(* IEC 61131-3 sources: TetherPLC/compat/tc3 (part 4) *)

(* ---- tc3_mcpath.st ---- *)
// Tc3_McCoordinatedMotion — MC path preparation + execution
// (TF5410 collision-avoidance / coordinated-motion bundle).
//
// This tranche implements the linear/dwell path subset:
//   MC_MoveLinearAbsolutePreparation, MC_MoveDirectPreparation
//   (flattened alias of the linear absolute segment),
//   MC_DwellTimePreparation, MC_MovePath.
// Path objects live in the tplc-path service via the FB_Path
// builtin; group membership comes from FB_McGroup.  Circular,
// blending and blocker segment types, MC_CalcTrafo, the CA move
// family, track following and compensation remain deferred.
//
// Flattened types (the ST dialect has no STRUCT/POINTER/REFERENCE
// support):
//   MC_PATH_DATA_REF     -> PathData : UDINT path handle (1..8)
//   Position (POINTER TO LREAL array) -> Position : ARRAY[0..15]
//                            OF LREAL + PositionCount
//   DwellTime (TIME)     -> DwellTime : UDINT milliseconds
//   BufferMode           -> UDINT (accepted, buffered queuing not
//                            modeled: every Execute edge appends a
//                            segment immediately)
//   AXES_GROUP_REF       -> AxesGroup : UDINT group handle
//
// Semantics:
//   * Preparation FBs append one segment on the Execute rising
//     edge. Linear segments store absolute user-unit positions and
//     trapezoid limits (Velocity/Acceleration; Deceleration and
//     Jerk are accepted but the service uses Acceleration for both
//     ramps). Dwell segments hold position for DwellTime ms.
//   * MC_MovePath on Execute captures each member axis's current
//     position (0x6064) as the path start, switches every member
//     to CSP mode (0x6060=8), then streams interpolated 0x607A
//     targets each scan until the path duration elapses. Positions
//     are interpolated in path parameter space on the dominant
//     axis, so all axes arrive together (coordinated motion).
//   * Segment targets chain: segment k starts where segment k-1
//     ended; the first segment starts at the captured positions.
//   * Busy stays TRUE while the path runs; Done pulses for one
//     scan at path end; Error carries service/axis failures.

// ---- shared path helper: ensure a valid PathData handle ----
// Returns TRUE and leaves `h` set to a usable path handle, or
// FALSE when the service table is full.

FUNCTION_BLOCK MC_MoveLinearAbsolutePreparation
VAR_INPUT
    Execute : BOOL;
    Position : ARRAY[0..15] OF LREAL;
    PositionCount : UDINT;
    Velocity : LREAL;
    Acceleration : LREAL;
    Deceleration : LREAL := 0.0;
    Jerk : LREAL := 0.0;
    BufferMode : UDINT := 1;
END_VAR
VAR_IN_OUT
    PathData : UDINT;
END_VAR
VAR_OUTPUT
    Error : BOOL;
    ErrorId : UDINT;
END_VAR
VAR
    p : FB_Path;
    exPrev : BOOL;
    edge : BOOL;
    i : UDINT;
END_VAR
edge := Execute AND NOT exPrev; exPrev := Execute;
Error := FALSE; ErrorId := 0;
IF edge THEN
    p.HANDLE := PathData;
    IF PathData = 0 THEN
        p.OP := 0; p();
        IF p.STATUS = 0 THEN PathData := p.HANDLE; END_IF;
    END_IF;
    IF PathData <> 0 AND PositionCount >= 1 AND
       PositionCount <= 16 THEN
        FOR i := 0 TO 15 DO p.POS[i] := Position[i]; END_FOR;
        p.OP := 2; p.AUX := 1; p.AUX2 := PositionCount;
        p.F1 := Velocity; p.F2 := Acceleration; p.F3 := 0.0;
        p.HANDLE := PathData; p();
        IF p.STATUS <> 0 THEN
            Error := TRUE;
            IF p.STATUS < 0 THEN ErrorId := 0 - p.STATUS; END_IF;
        END_IF;
    ELSE
        Error := TRUE; ErrorId := 16#4D01;
    END_IF;
END_IF;
END_FUNCTION_BLOCK

// MC_MoveDirectPreparation: TwinCAT "direct" segments are absolute
// linear moves without blending lookahead.  Flattened to the same
// linear segment; BufferMode is accepted for signature parity.
FUNCTION_BLOCK MC_MoveDirectPreparation
VAR_INPUT
    Execute : BOOL;
    Position : ARRAY[0..15] OF LREAL;
    PositionCount : UDINT;
    Velocity : LREAL;
    Acceleration : LREAL;
    Deceleration : LREAL := 0.0;
    Jerk : LREAL := 0.0;
    BufferMode : UDINT := 1;
END_VAR
VAR_IN_OUT
    PathData : UDINT;
END_VAR
VAR_OUTPUT
    Error : BOOL;
    ErrorId : UDINT;
END_VAR
VAR
    p : FB_Path;
    exPrev : BOOL;
    edge : BOOL;
    i : UDINT;
END_VAR
edge := Execute AND NOT exPrev; exPrev := Execute;
Error := FALSE; ErrorId := 0;
IF edge THEN
    p.HANDLE := PathData;
    IF PathData = 0 THEN
        p.OP := 0; p();
        IF p.STATUS = 0 THEN PathData := p.HANDLE; END_IF;
    END_IF;
    IF PathData <> 0 AND PositionCount >= 1 AND
       PositionCount <= 16 THEN
        FOR i := 0 TO 15 DO p.POS[i] := Position[i]; END_FOR;
        p.OP := 2; p.AUX := 1; p.AUX2 := PositionCount;
        p.F1 := Velocity; p.F2 := Acceleration; p.F3 := 0.0;
        p.HANDLE := PathData; p();
        IF p.STATUS <> 0 THEN
            Error := TRUE;
            IF p.STATUS < 0 THEN ErrorId := 0 - p.STATUS; END_IF;
        END_IF;
    ELSE
        Error := TRUE; ErrorId := 16#4D01;
    END_IF;
END_IF;
END_FUNCTION_BLOCK

FUNCTION_BLOCK MC_DwellTimePreparation
VAR_INPUT
    Execute : BOOL;
    DwellTime : UDINT;   // milliseconds (TIME flattened)
    BufferMode : UDINT := 1;
END_VAR
VAR_IN_OUT
    PathData : UDINT;
END_VAR
VAR_OUTPUT
    Error : BOOL;
    ErrorId : UDINT;
END_VAR
VAR
    p : FB_Path;
    exPrev : BOOL;
    edge : BOOL;
END_VAR
edge := Execute AND NOT exPrev; exPrev := Execute;
Error := FALSE; ErrorId := 0;
IF edge THEN
    p.HANDLE := PathData;
    IF PathData = 0 THEN
        p.OP := 0; p();
        IF p.STATUS = 0 THEN PathData := p.HANDLE; END_IF;
    END_IF;
    IF PathData <> 0 THEN
        p.OP := 2; p.AUX := 3; p.AUX2 := 0;
        p.F1 := 0.0; p.F2 := 0.0; p.F3 := DwellTime;
        p.HANDLE := PathData; p();
        IF p.STATUS <> 0 THEN
            Error := TRUE;
            IF p.STATUS < 0 THEN ErrorId := 0 - p.STATUS; END_IF;
        END_IF;
    ELSE
        Error := TRUE; ErrorId := 16#4D01;
    END_IF;
END_IF;
END_FUNCTION_BLOCK

FUNCTION_BLOCK MC_MovePath
VAR_INPUT
    Execute : BOOL;
END_VAR
VAR_IN_OUT
    AxesGroup : UDINT;
    PathData : UDINT;
END_VAR
VAR_OUTPUT
    Done : BOOL;
    Busy : BOOL;
    CommandAborted : BOOL;
    Error : BOOL;
    ErrorId : UDINT;
END_VAR
VAR
    mg : FB_McGroup;
    p : FB_Path;
    ax : FB_MotionAxis;
    exPrev : BOOL;
    exEdge : BOOL;
    active : BOOL;
    issued : BOOL;
    t0 : LREAL;
    pathT : LREAL;
    lastNow : LREAL;
    blkWait : BOOL;
    trafoGen : UDINT;
    lastTrafoGen : UDINT;
    dn : LREAL;
    i : UDINT;
    n : UDINT;
    axh : UDINT;
    startPos : ARRAY[0..15] OF LREAL;
END_VAR
mg.GRP := AxesGroup;
mg.OP := 10; mg();
AxesGroup := mg.GRP;
n := mg.NAXES;
exEdge := Execute AND NOT exPrev; exPrev := Execute;
Done := FALSE; Busy := FALSE;
CommandAborted := FALSE; Error := FALSE; ErrorId := 0;
IF exEdge THEN
    active := TRUE; issued := FALSE;
END_IF;
IF active THEN
    IF NOT issued THEN
        /* capture current positions as the path start */
        FOR i := 0 TO 15 DO
            startPos[i] := 0.0;
            IF i < n THEN
                axh := mg.AXES[i];
                ax.AXIS := axh; ax.OP := 4; ax.INDEX := 16#6064; ax();
                startPos[i] := DINT_TO_LREAL(ax.VALUE);
            END_IF;
        END_FOR;
        FOR i := 0 TO 15 DO p.POS[i] := startPos[i]; END_FOR;
        p.OP := 3; p.AUX := n; p.HANDLE := PathData; p();
        IF p.STATUS <> 0 THEN
            Error := TRUE;
            IF p.STATUS < 0 THEN ErrorId := 0 - p.STATUS; END_IF;
            active := FALSE;
        ELSE
            PathData := p.HANDLE;
            /* bind the path to the group for trajectory readback */
            p.OP := 9; p.AUX := AxesGroup; p.HANDLE := PathData; p();
            t0 := p.NOW;
            pathT := 0.0; lastNow := p.NOW;
            /* switch members to CSP mode for 0x607A streaming */
            FOR i := 0 TO 15 DO
                IF i < n THEN
                    axh := mg.AXES[i];
                    ax.AXIS := axh; ax.OP := 5;
                    ax.INDEX := 16#6060; ax.VALUE := 8; ax();
                END_IF;
            END_FOR;
            issued := TRUE;
        END_IF;
    END_IF;
    IF issued THEN
        /* blocker query freezes path time while the path is held
           at an unreleased blocker gate */
        p.OP := 7; p.HANDLE := PathData; p();
        blkWait := p.AUX = 1;
        dn := p.NOW - lastNow; lastNow := p.NOW;
        IF NOT blkWait THEN pathT := pathT + dn; END_IF;
        /* apply pending coordinate-transform markers: the service
           bumps AUX2 whenever the pending id changes */
        p.OP := 11; p.HANDLE := PathData; p();
        trafoGen := p.AUX2;
        IF trafoGen <> lastTrafoGen AND p.F1 <> 0.0 THEN
            lastTrafoGen := trafoGen;
            mg.OP := 9; mg.COORD := LREAL_TO_DINT(p.F1); mg();
        END_IF;
        p.OP := 4; p.F1 := pathT; p.HANDLE := PathData; p();
        IF p.STATUS <> 0 THEN
            Error := TRUE;
            IF p.STATUS < 0 THEN ErrorId := 0 - p.STATUS; END_IF;
            active := FALSE; CommandAborted := TRUE;
        ELSE
            FOR i := 0 TO 15 DO
                IF i < n THEN
                    axh := mg.AXES[i];
                    ax.AXIS := axh; ax.OP := 5;
                    ax.INDEX := 16#607A;
                    ax.VALUE := LREAL_TO_DINT(p.POS[i]); ax();
                END_IF;
            END_FOR;
            IF p.DONE = 1 THEN
                Done := TRUE; active := FALSE;
            END_IF;
        END_IF;
    END_IF;
    Busy := active;
END_IF;
END_FUNCTION_BLOCK

// MC_MoveCircularAbsolutePreparation: appends a circular segment.
// CircMode flattens MC_CIRC_MODE (1=mcCircModeCenter: AuxPoint is
// the circle center and must be equidistant from start/end;
// 2=mcCircModeBorder: AuxPoint lies on the circle). The circle is
// evaluated in the plane of position entries 0/1; entries >=2
// interpolate linearly. PathChoice: 1=counter-clockwise,
// 2=clockwise. TransitionMode/TransitionParameter/InvokeId/
// DynamicConstraints are accepted for signature parity but not
// modeled.
FUNCTION_BLOCK MC_MoveCircularAbsolutePreparation
VAR_INPUT
    Execute : BOOL;
    CircMode : UDINT;
    AuxPoint : ARRAY[0..15] OF LREAL;
    AuxPointCount : UDINT;
    EndPoint : ARRAY[0..15] OF LREAL;
    EndPointCount : UDINT;
    PathChoice : UDINT := 1;
    Velocity : LREAL;
    Acceleration : LREAL;
    Deceleration : LREAL := 0.0;
    Jerk : LREAL := 0.0;
    BufferMode : UDINT := 1;
    TransitionMode : UDINT := 0;
    TransitionParameter : ARRAY[0..15] OF LREAL;
    TransitionParameterCount : UDINT := 0;
    InvokeId : UDINT := 0;
END_VAR
VAR_IN_OUT
    PathData : UDINT;
END_VAR
VAR_OUTPUT
    Error : BOOL;
    ErrorId : UDINT;
END_VAR
VAR
    p : FB_Path;
    exPrev : BOOL;
    edge : BOOL;
    i : UDINT;
END_VAR
edge := Execute AND NOT exPrev; exPrev := Execute;
Error := FALSE; ErrorId := 0;
IF edge THEN
    p.HANDLE := PathData;
    IF PathData = 0 THEN
        p.OP := 0; p();
        IF p.STATUS = 0 THEN PathData := p.HANDLE; END_IF;
    END_IF;
    IF PathData <> 0 AND EndPointCount >= 1 AND EndPointCount <= 16
       AND CircMode >= 1 AND CircMode <= 2 THEN
        FOR i := 0 TO 15 DO
            p.POS[i] := EndPoint[i];
            p.AUXP[i] := AuxPoint[i];
        END_FOR;
        p.OP := 6; p.AUX := CircMode; p.FLAGS := AuxPointCount;
        p.AUX2 := EndPointCount; p.F3 := PathChoice;
        p.F1 := Velocity; p.F2 := Acceleration;
        p.HANDLE := PathData; p();
        IF p.STATUS <> 0 THEN
            Error := TRUE;
            IF p.STATUS < 0 THEN ErrorId := 0 - p.STATUS; END_IF;
        END_IF;
    ELSE
        Error := TRUE; ErrorId := 16#4D01;
    END_IF;
END_IF;
END_FUNCTION_BLOCK

// MC_MoveBlendingPreparation: appends a junction transition segment.
// TwinCAT uses it to program velocity blending between segments;
// this implementation holds the path end position for
// TransitionParameter[0] milliseconds (real corner-cutting/lookahead
// blending is not modeled — documented deviation). Velocity/
// Acceleration/Deceleration/Jerk are accepted for signature parity.
FUNCTION_BLOCK MC_MoveBlendingPreparation
VAR_INPUT
    Execute : BOOL;
    Velocity : LREAL;
    Acceleration : LREAL;
    Deceleration : LREAL := 0.0;
    Jerk : LREAL := 0.0;
    BufferMode : UDINT := 1;
    TransitionMode : UDINT := 0;
    TransitionParameter : ARRAY[0..15] OF LREAL;
    TransitionParameterCount : UDINT := 0;
    InvokeId : UDINT := 0;
END_VAR
VAR_IN_OUT
    PathData : UDINT;
END_VAR
VAR_OUTPUT
    Error : BOOL;
    ErrorId : UDINT;
END_VAR
VAR
    p : FB_Path;
    exPrev : BOOL;
    edge : BOOL;
END_VAR
edge := Execute AND NOT exPrev; exPrev := Execute;
Error := FALSE; ErrorId := 0;
IF edge THEN
    p.HANDLE := PathData;
    IF PathData = 0 THEN
        p.OP := 0; p();
        IF p.STATUS = 0 THEN PathData := p.HANDLE; END_IF;
    END_IF;
    IF PathData <> 0 THEN
        p.OP := 2; p.AUX := 4; p.AUX2 := 0;
        p.F1 := 0.0; p.F2 := 0.0;
        IF TransitionParameterCount >= 1 THEN
            p.F3 := TransitionParameter[0];
        ELSE
            p.F3 := 0.0;
        END_IF;
        p.HANDLE := PathData; p();
        IF p.STATUS <> 0 THEN
            Error := TRUE;
            IF p.STATUS < 0 THEN ErrorId := 0 - p.STATUS; END_IF;
        END_IF;
    ELSE
        Error := TRUE; ErrorId := 16#4D01;
    END_IF;
END_IF;
END_FUNCTION_BLOCK

// MC_BlockerPreparation: appends a blocker gate at the current path
// junction. The path holds position there during MC_MovePath until
// MC_ReleaseBlocker opens the gate. BufferMode is accepted for
// signature parity.
FUNCTION_BLOCK MC_BlockerPreparation
VAR_INPUT
    Execute : BOOL;
    BlockerId : UDINT;
    BufferMode : UDINT := 1;
END_VAR
VAR_IN_OUT
    PathData : UDINT;
END_VAR
VAR_OUTPUT
    Error : BOOL;
    ErrorId : UDINT;
END_VAR
VAR
    p : FB_Path;
    exPrev : BOOL;
    edge : BOOL;
END_VAR
edge := Execute AND NOT exPrev; exPrev := Execute;
Error := FALSE; ErrorId := 0;
IF edge THEN
    p.HANDLE := PathData;
    IF PathData = 0 THEN
        p.OP := 0; p();
        IF p.STATUS = 0 THEN PathData := p.HANDLE; END_IF;
    END_IF;
    IF PathData <> 0 AND BlockerId > 0 THEN
        p.OP := 2; p.AUX := 5; p.AUX2 := 0;
        p.F1 := 0.0; p.F2 := 0.0; p.F3 := BlockerId;
        p.HANDLE := PathData; p();
        IF p.STATUS <> 0 THEN
            Error := TRUE;
            IF p.STATUS < 0 THEN ErrorId := 0 - p.STATUS; END_IF;
        END_IF;
    ELSE
        Error := TRUE; ErrorId := 16#4D01;
    END_IF;
END_IF;
END_FUNCTION_BLOCK

// MC_ReleaseBlocker: opens every blocker gate with the given id on
// the next eval. The TwinCAT signature carries only AxesGroup; the
// flattened implementation releases by BlockerId across all path
// objects (blocker ids are user-unique per machine).
FUNCTION_BLOCK MC_ReleaseBlocker
VAR_INPUT
    Execute : BOOL;
    BlockerId : UDINT;
END_VAR
VAR_IN_OUT
    AxesGroup : UDINT;
END_VAR
VAR_OUTPUT
    Done : BOOL;
    Busy : BOOL;
    Error : BOOL;
    ErrorId : UDINT;
END_VAR
VAR
    p : FB_Path;
    mg : FB_McGroup;
    exPrev : BOOL;
    edge : BOOL;
    ok : BOOL;
END_VAR
ok := FALSE;
edge := Execute AND NOT exPrev;
mg.GRP := AxesGroup; mg.OP := 1; mg();
AxesGroup := mg.GRP;
IF edge THEN
    p.OP := 8; p.F1 := BlockerId; p();
    IF p.STATUS = 0 THEN ok := TRUE; END_IF;
END_IF;
exPrev := Execute;
Done := ok; Busy := FALSE;
Error := edge AND NOT ok;
IF edge AND p.STATUS < 0 THEN ErrorId := 0 - p.STATUS; END_IF;
END_FUNCTION_BLOCK

// MC_GroupReadBlockerStatus: reports whether the most recent path
// eval is held at an unreleased blocker. The group linkage is
// approximated — the service reports the last-evaluated path's gate
// state.
FUNCTION_BLOCK MC_GroupReadBlockerStatus
VAR_INPUT
    Enable : BOOL;
END_VAR
VAR_IN_OUT
    AxesGroup : UDINT;
END_VAR
VAR_OUTPUT
    Valid : BOOL;
    Busy : BOOL;
    Blocked : BOOL;
    BlockerId : UDINT;
    Error : BOOL;
    ErrorId : UDINT;
END_VAR
VAR
    p : FB_Path;
    mg : FB_McGroup;
END_VAR
Valid := FALSE; Busy := FALSE; Blocked := FALSE;
BlockerId := 0; Error := FALSE; ErrorId := 0;
mg.GRP := AxesGroup; mg.OP := 6; mg();
IF Enable AND mg.STATUS = 0 THEN
    Valid := TRUE;
    p.OP := 7; p();
    IF p.STATUS = 0 THEN
        Blocked := p.AUX = 1;
        BlockerId := LREAL_TO_DINT(p.F1);
    ELSE
        Error := TRUE;
        IF p.STATUS < 0 THEN ErrorId := 0 - p.STATUS; END_IF;
    END_IF;
END_IF;
END_FUNCTION_BLOCK

// MC_GroupReadTrajectoryInformation: reads the current and next
// path segments for the group the executing MC_MovePath is bound
// to. Entries flatten MC_TRAJECTORY_ENTRY: InvokeId is approximated
// by the 1-based segment index, Active marks blend/blocker
// segments, RemainingDuration is seconds and
// RemainingCartesianLength is dominant-axis user units, all as of
// the most recent path eval.
FUNCTION_BLOCK MC_GroupReadTrajectoryInformation
VAR_INPUT
    Enable : BOOL;
END_VAR
VAR_IN_OUT
    AxesGroup : UDINT;
END_VAR
VAR_OUTPUT
    Valid : BOOL;
    Busy : BOOL;
    Error : BOOL;
    ErrorId : UDINT;
    EntryCount : UDINT;
    TrajInvokeId : ARRAY[0..9] OF UDINT;
    TrajActive : ARRAY[0..9] OF BOOL;
    TrajRemLen : ARRAY[0..9] OF LREAL;
    TrajRemDur : ARRAY[0..9] OF LREAL;
END_VAR
VAR
    p : FB_Path;
    mg : FB_McGroup;
    i : UDINT;
END_VAR
Valid := FALSE; Busy := FALSE; Error := FALSE; ErrorId := 0;
EntryCount := 0;
mg.GRP := AxesGroup; mg.OP := 6; mg();
IF Enable AND mg.STATUS = 0 THEN
    Valid := TRUE;
    p.OP := 10; p.AUX := AxesGroup; p();
    IF p.STATUS = 0 THEN
        EntryCount := p.NSEG;
        FOR i := 0 TO 9 DO
            TrajInvokeId[i] := p.TRID[i];
            TrajActive[i] := p.TACT[i] = 1;
            TrajRemLen[i] := p.AUXP[i];
            TrajRemDur[i] := p.POS[i];
        END_FOR;
    ELSE
        Error := TRUE;
        IF p.STATUS < 0 THEN ErrorId := 0 - p.STATUS; END_IF;
    END_IF;
END_IF;
END_FUNCTION_BLOCK

// MC_SetCoordinateTransformPreparation: inserts a reference-system
// change marker into the path (TwinCAT signature has no Execute;
// the flattened version appends when the CoordTransform input
// changes value). MC_MovePath applies the group's coordinate
// transform when path time reaches the marker.
FUNCTION_BLOCK MC_SetCoordinateTransformPreparation
VAR_INPUT
    PathData : UDINT;
    CoordTransform : UDINT;
END_VAR
VAR_OUTPUT
    Error : BOOL;
    ErrorId : UDINT;
END_VAR
VAR
    p : FB_Path;
    prevCoord : UDINT := 0;
END_VAR
Error := FALSE; ErrorId := 0;
IF CoordTransform <> prevCoord AND CoordTransform <> 0 THEN
    p.HANDLE := PathData;
    IF PathData <> 0 THEN
        p.OP := 2; p.AUX := 6; p.AUX2 := 0;
        p.F1 := 0.0; p.F2 := 0.0; p.F3 := CoordTransform;
        p.HANDLE := PathData; p();
        IF p.STATUS <> 0 THEN
            Error := TRUE;
            IF p.STATUS < 0 THEN ErrorId := 0 - p.STATUS; END_IF;
        END_IF;
    ELSE
        Error := TRUE; ErrorId := 16#4D01;
    END_IF;
END_IF;
prevCoord := CoordTransform;
END_FUNCTION_BLOCK

(* ---- tc3_mll.st ---- *)
// tc3_mll.st — Tc3_MLL surface (TF38x0): ML inference prediction
// block.  TwinCAT loads an ONNX/TF-lite model into the ML runtime
// and runs async predictions.  TetherPLC ships no inference
// engine, so the default path is honest engine-absent: commands
// are accepted, Busy runs a bounded handshake, then Error with
// ErrorId=1 (engine-unavailable) — predictions are never faked.
//
// A pure-ST simulation mode is provided for logic testing:
// with UseSimulation=TRUE the block runs a deterministic
// single-output linear model  y = SUM(Wi * Xi) + Bias  over the
// caller-supplied weights — no engine required, and the result is
// honest arithmetic, not a canned answer.
//
// Differences from the TwinCAT FB (docs/plc/compat/README.md):
//   - stPredictionParameter is decomposed into plain inputs
//     (ModelPath, InputCount, X0..X7, UseSimulation, W0..W7, Bias);
//     TetherPLC has no struct/method surface in compat ST.
//   - CheckPreferredIODataTypes is exposed as inputs
//     FmtIn/FmtOut + output FmtPreferred (Tc float32/int32 codes:
//     1=f32, 2=i32, 3=i64, 4=f64 — preferred set {1,2}).
//   - ipResultMessage / I_TcMessage is replaced by UDINT ErrorId:
//     0 none, 1 engine-unavailable, 2 bad-input-rank,
//     3 bad-model, 4 sim-dtype-mismatch, 5 aborted.
//   - Predictions expose a scalar Y plus valid flag; the real
//     tensor output surface needs the engine.

// ---- FB_MllPrediction (TwinCAT §6.2.2.1) ----
FUNCTION_BLOCK FB_MllPrediction
VAR_INPUT
    Execute : BOOL;             // rising edge starts a prediction
    Abort : BOOL;
    ModelPath : STRING;         // ONNX model path (engine mode)
    InputCount : UDINT;         // active X lanes, 1..8
    UseSimulation : BOOL;       // TRUE: run the built-in linear sim
    X0 : LREAL; X1 : LREAL; X2 : LREAL; X3 : LREAL;
    X4 : LREAL; X5 : LREAL; X6 : LREAL; X7 : LREAL;
    W0 : LREAL; W1 : LREAL; W2 : LREAL; W3 : LREAL;
    W4 : LREAL; W5 : LREAL; W6 : LREAL; W7 : LREAL;
    Bias : LREAL;
    FmtIn : UDINT;              // CheckPreferredIODataTypes surface
    FmtOut : UDINT;
END_VAR
VAR_OUTPUT
    Busy : BOOL;
    Error : BOOL;
    ErrorId : UDINT;
    Done : BOOL;
    Y : LREAL;                  // prediction (simulation mode)
    YValid : BOOL;
    FmtPreferred : BOOL;
END_VAR
VAR
    phase : INT;                 // 0 idle, 1 handshake, 2 done
    tmo : UDINT;
    acc : LREAL;
    lanes : UDINT;
END_VAR
    Done := FALSE;
    YValid := FALSE;

    // preferred-IO-type check: TCML supports f32/i32 natively
    FmtPreferred := ((FmtIn = 1) OR (FmtIn = 2)) AND
                    ((FmtOut = 1) OR (FmtOut = 2));

    IF phase = 0 THEN
        Busy := FALSE;
        IF Execute THEN
            Busy := TRUE;
            Error := FALSE;
            ErrorId := 0;
            Y := 0.0;
            tmo := 0;
            // parameter validation first (mirrors TwinCAT checks)
            IF InputCount = 0 OR InputCount > 8 THEN
                Error := TRUE;
                ErrorId := 2;        // bad-input-rank
                phase := 2;
            ELSIF NOT UseSimulation AND ModelPath = '' THEN
                Error := TRUE;
                ErrorId := 3;        // bad-model: no path, no engine
                phase := 2;
            ELSIF UseSimulation THEN
                // deterministic linear inference: y = W.x + Bias
                acc := Bias;
                lanes := InputCount;
                IF lanes > 0 THEN acc := acc + W0 * X0; END_IF;
                IF lanes > 1 THEN acc := acc + W1 * X1; END_IF;
                IF lanes > 2 THEN acc := acc + W2 * X2; END_IF;
                IF lanes > 3 THEN acc := acc + W3 * X3; END_IF;
                IF lanes > 4 THEN acc := acc + W4 * X4; END_IF;
                IF lanes > 5 THEN acc := acc + W5 * X5; END_IF;
                IF lanes > 6 THEN acc := acc + W6 * X6; END_IF;
                IF lanes > 7 THEN acc := acc + W7 * X7; END_IF;
                Y := acc;
                YValid := TRUE;
                Busy := FALSE;
                phase := 2;
            ELSE
                phase := 1;          // engine handshake window
            END_IF;
        END_IF;
    ELSIF phase = 1 THEN
        tmo := tmo + 1;
        IF tmo >= 4 THEN
            Busy := FALSE;
            Error := TRUE;
            ErrorId := 1;            // engine-unavailable
            phase := 2;
        END_IF;
    ELSE
        Busy := FALSE;
        IF NOT Execute THEN
            phase := 0;              // re-arm on falling edge
        END_IF;
    END_IF;

    IF Abort AND phase = 1 THEN
        Busy := FALSE;
        Error := TRUE;
        ErrorId := 5;
        phase := 2;
    END_IF;
    Done := (phase = 2);
END_FUNCTION_BLOCK

(* ---- tc3_nccam.st ---- *)
// tc3_nccam.st — TF5050 Tc3_NC_Camming compatibility surface.
//
// Electronic camming couples a slave axis to a master axis through
// a cam table (master position -> slave position).  TwinCAT models
// this as MC_CAM_REF table objects shared between the motion-
// function FBs (MC_WriteMotionFunction*) and the coupling FBs
// (MC_CamTableSelect/MC_CamIn/MC_CamOut/MC_CamAdd/...).  This
// dialect has no REFERENCE TO, so the table lives inside the
// coupling FB as public member arrays MasterPosT/SlavePosT
// (LREAL, sorted ascending by master position, up to 64 points) —
// the documented flattening of MC_CAM_REF.  Points can also be
// written through the Pt* edge inputs (the
// MC_WriteMotionFunctionPoint shape).
//
// FB_McCamAxis (builtin FB_MotionAxis) supplies the axis handles:
// MasterAxis/SlaveAxis are the UDINT handles returned by
// FB_MotionAxis OP=1 create — the same AXIS_REF flattening used by
// compat/tc2/tc2_mc2.st.
//
// Semantics: while Execute is TRUE the FB polls both axes, reads
// the master position actual (0x6064), applies
//   mt = masterActual * MasterScaling + MasterOffset
// looks the cam table up (linear interpolation, clamped ends,
// optional periodic wrap), applies
//   st = slaveTablePos * SlaveScaling + SlaveOffset
// and writes the slave position target (0x607A) every scan.  The
// slave axis must be powered and in CSP mode (the case/program
// sets 0x6060=8 once; the FB does not change modes).  Invert=TRUE
// swaps the coupling direction (MC_CamIn vs MC_CamOut roles).
//
// Mapping notes (documented deviations):
//   - MC_CamAdd/Exchange/Remove multi-plate blending, online
//     change modes, cam-table file I/O, slave-dynamics and
//     characteristics reads are not implemented; single-table
//     linear coupling only.
//   - LREAL engineering units map onto the backend's int32 user
//     units at the axis boundary (same documented gap as tc2_mc2).
//
// SPDX-License-Identifier: Apache-2.0 OR MPL-2.0

FUNCTION_BLOCK FB_McCamCoupling
VAR_INPUT
    Execute : BOOL;              // coupling active while TRUE
    MasterAxis : UDINT;          // FB_MotionAxis handle
    SlaveAxis : UDINT;           // FB_MotionAxis handle
    Periodic : BOOL;             // wrap master position
    Invert : BOOL;               // swap master/slave roles
    CamTableID : UDINT;          // echoed on CamTableID output
    MasterOffset : LREAL := 0.0;
    SlaveOffset : LREAL := 0.0;
    MasterScaling : LREAL := 1.0;
    SlaveScaling : LREAL := 1.0;
    // MC_WriteMotionFunctionPoint shape (edge writes one point)
    WritePt : BOOL;
    PtIndex : UDINT;             // 0..63
    PtMaster : LREAL;
    PtSlave : LREAL;
    ClearTable : BOOL;           // edge: TableCount := 0
END_VAR
VAR_OUTPUT
    Done : BOOL;
    Busy : BOOL;
    Error : BOOL;
    ErrorID : UDINT;
    InSync : BOOL;
    CamTableIDOut : UDINT;
    CamSlavePos : LREAL;         // last interpolated slave pos
    TableCountOut : UDINT;
END_VAR
VAR
    axM : FB_MotionAxis;
    axS : FB_MotionAxis;
    prevExec : BOOL;
    prevWr : BOOL;
    prevClr : BOOL;
    i : UDINT;
    mt : LREAL;
    st : LREAL;
    frac : LREAL;
    range : LREAL;
    wraps : UDINT;
    masterH : UDINT;
    slaveH : UDINT;
    mActual : DINT;
    seg : UDINT;
    found : BOOL;
    // public table storage (MC_CAM_REF flattening)
    MasterPosT : ARRAY[0..63] OF LREAL;
    SlavePosT : ARRAY[0..63] OF LREAL;
    TableCount : UDINT;
END_VAR
    Busy := FALSE;
    Error := FALSE;
    ErrorID := 0;
    CamTableIDOut := CamTableID;
    TableCountOut := TableCount;

    // table maintenance edges
    IF ClearTable AND NOT prevClr THEN
        TableCount := 0;
    END_IF;
    IF WritePt AND NOT prevWr AND PtIndex < 64 THEN
        MasterPosT[PtIndex] := PtMaster;
        SlavePosT[PtIndex] := PtSlave;
        IF PtIndex >= TableCount THEN
            TableCount := PtIndex + 1;
        END_IF;
    END_IF;
    prevWr := WritePt;
    prevClr := ClearTable;

    masterH := MasterAxis;
    slaveH := SlaveAxis;
    IF Invert THEN
        masterH := SlaveAxis;
        slaveH := MasterAxis;
    END_IF;

    IF Execute THEN
        // advance dynamics once per scan on both axes
        axM.AXIS := masterH; axM.OP := 3; axM();
        axS.AXIS := slaveH;   axS.OP := 3; axS();

        IF axM.STATUS < 0 OR axS.STATUS < 0 THEN
            Error := TRUE;
            ErrorID := 1;
        ELSIF TableCount < 2 THEN
            // need at least two points for interpolation
            InSync := FALSE;
        ELSE
            // master position actual -> scaled table coordinate
            axM.OP := 6; axM();
            mActual := axM.POS_ACTUAL;
            mt := DINT_TO_LREAL(mActual) * MasterScaling + MasterOffset;

            // locate segment (table sorted ascending by master pos)
            seg := 0;
            found := FALSE;
            FOR i := 0 TO TableCount - 2 DO
                IF mt <= MasterPosT[i + 1] THEN
                    seg := i;
                    found := TRUE;
                END_IF;
            END_FOR;
            IF mt < MasterPosT[0] THEN
                st := SlavePosT[0];
            ELSIF mt > MasterPosT[TableCount - 1] THEN
                IF Periodic AND
                   MasterPosT[TableCount - 1] > MasterPosT[0] THEN
                    range := MasterPosT[TableCount - 1] - MasterPosT[0];
                    wraps := 0;
                    WHILE mt > MasterPosT[TableCount - 1] AND wraps < 1024 DO
                        mt := mt - range;
                        wraps := wraps + 1;
                    END_WHILE;
                    // re-locate after wrap
                    FOR i := 0 TO TableCount - 2 DO
                        IF mt <= MasterPosT[i + 1] THEN
                            seg := i;
                            found := TRUE;
                        END_IF;
                    END_FOR;
                    IF found AND MasterPosT[seg + 1] > MasterPosT[seg] THEN
                        frac := (mt - MasterPosT[seg]) /
                                (MasterPosT[seg + 1] - MasterPosT[seg]);
                        st := SlavePosT[seg] +
                              frac * (SlavePosT[seg + 1] - SlavePosT[seg]);
                    ELSE
                        st := SlavePosT[TableCount - 1];
                    END_IF;
                ELSE
                    st := SlavePosT[TableCount - 1];
                END_IF;
            ELSIF NOT found THEN
                st := SlavePosT[TableCount - 1];
            ELSE
                IF MasterPosT[seg + 1] > MasterPosT[seg] THEN
                    frac := (mt - MasterPosT[seg]) /
                            (MasterPosT[seg + 1] - MasterPosT[seg]);
                    st := SlavePosT[seg] +
                          frac * (SlavePosT[seg + 1] - SlavePosT[seg]);
                ELSE
                    st := SlavePosT[seg];
                END_IF;
            END_IF;

            // slave target in backend units
            st := st * SlaveScaling + SlaveOffset;
            CamSlavePos := st;
            axS.OP := 5;
            axS.INDEX := 16#607A;
            axS.VALUE := LREAL_TO_DINT(st);
            axS();
            IF axS.STATUS < 0 THEN
                Error := TRUE;
                ErrorID := 2;
            END_IF;
            InSync := NOT Error;
        END_IF;
        Done := Execute;
    ELSE
        InSync := FALSE;
        Done := FALSE;
        CamSlavePos := 0.0;
    END_IF;
    prevExec := Execute;
END_FUNCTION_BLOCK

(* ---- tc3_pjlink.st ---- *)
// Tc3_PJLink -> JBMIA PJLink projector client wrappers.
// TwinCAT's FB_PJLink is an auto-managed connection object with
// EventLogger events and AMS NetID routing; TetherPLC adapts it
// to the poll-driven service model used by the other compat
// libraries (one transaction per EXEC edge, service-enforced
// timeout, connect-per-command).
// Differences from the TwinCAT FB, documented in
// docs/plc/compat/README.md:
//   - No persistent keep-alive session, no tStatusUpdateTime
//     polling, no sServerNetID routing (direct IPv4 only),
//     no I_TcMessage/HRESULT/EventLogger surfaces.
//   - PASSWORD drives the PJLink digest exchange automatically
//     when the projector greets `PJLINK 1 <nonce>`.
//   - PJLink "class" is the digit after '%' (standard commands
//     use class 1); nCmd is the 4-char body ("POWR","INPT",
//     "AVMT","ERST","INFO","NAME","INFM","LAMP", ...).
//   - nStatus mirrors TplcPjlinkRespInfo: 0=pending 1=ok
//     2=timeout 3=error 4=badresp 5=authfail. PJLink-level
//     command errors arrive as sValue="ERR<n>" with nStatus=1.
// Sources: docs/plc/plan/21-twincat-libraries.md (TF8020 PJLink).

FUNCTION_BLOCK FB_PJLink
VAR_INPUT
    sHost : STRING[15];          // dotted-quad projector IPv4
    nPort : UDINT := 4352;       // 0 = 4352
    nCls : UDINT := 1;           // PJLink class digit 0..9
    sCmd : STRING[4];            // 4-char command body
    sParam : STRING[128];        // "?" for queries
    sPassword : STRING[32];      // "" = no auth
    bExecute : BOOL;
    tTimeout : TIME := T#2S;
END_VAR
VAR_OUTPUT
    bBusy : BOOL;
    bDone : BOOL;
    bError : BOOL;
    nErrId : UDINT;
    nStatus : DINT;
    bAuthed : BOOL;
    nRespCls : UDINT;
    nRespCmd : UDINT;            // 4-char body packed BE ASCII
    nValueLen : UDINT;           // full value length
    sValue : STRING[127];        // response value text
END_VAR
VAR
    pjl : FB_Pjlink;
END_VAR
    pjl.HOST := sHost;
    pjl.PORT := nPort;
    pjl.CLS := nCls;
    pjl.CMD := sCmd;
    pjl.PARAM := sParam;
    pjl.PASSWORD := sPassword;
    pjl.TIMEOUT := tTimeout;
    pjl.EXEC := bExecute;
    pjl();
    bBusy := pjl.BUSY;
    bDone := pjl.DONE;
    nStatus := pjl.STATUS;
    nErrId := pjl.ERRID;
    bAuthed := pjl.AUTHED;
    nRespCls := pjl.R_CLS;
    nRespCmd := pjl.R_CMD;
    nValueLen := pjl.R_VLEN;
    sValue := pjl.R_VALUE;
    bError := (pjl.ERRID <> 0) OR (pjl.STATUS >= 2);
END_FUNCTION_BLOCK

// Power on/off/query — TwinCAT PowerOn/PowerOff methods folded
// into one poll-model FB. nMode: 0=off 1=on 2=query.
FUNCTION_BLOCK FB_PJLink_Power
VAR_INPUT
    sHost : STRING[15];
    nPort : UDINT := 4352;
    sPassword : STRING[32] := '';
    nMode : UDINT;               // 0=off 1=on 2=query
    bExecute : BOOL;
    tTimeout : TIME := T#2S;
END_VAR
VAR_OUTPUT
    bBusy : BOOL;
    bDone : BOOL;
    bError : BOOL;
    nErrId : UDINT;
    nStatus : DINT;
    bAuthed : BOOL;
    sValue : STRING[127];        // query: "0".."3" power state
END_VAR
VAR
    pjl : FB_PJLink;
END_VAR
    pjl.sHost := sHost;
    pjl.nPort := nPort;
    pjl.nCls := 1;
    pjl.sCmd := 'POWR';
    IF nMode = 2 THEN
        pjl.sParam := '?';
    ELSIF nMode = 1 THEN
        pjl.sParam := '1';
    ELSE
        pjl.sParam := '0';
    END_IF;
    pjl.sPassword := sPassword;
    pjl.tTimeout := tTimeout;
    pjl.bExecute := bExecute;
    pjl();
    bBusy := pjl.bBusy;
    bDone := pjl.bDone;
    bError := pjl.bError;
    nErrId := pjl.nErrId;
    nStatus := pjl.nStatus;
    bAuthed := pjl.bAuthed;
    sValue := pjl.sValue;
END_FUNCTION_BLOCK

// Input select/query — TwinCAT SetInputType/SetInputChannel
// methods. nMode: 0=set (sParam = input number, e.g. "31")
// 1=query.
FUNCTION_BLOCK FB_PJLink_Input
VAR_INPUT
    sHost : STRING[15];
    nPort : UDINT := 4352;
    sPassword : STRING[32] := '';
    nMode : UDINT;               // 0=set 1=query
    sInput : STRING[8];          // input number when nMode=0
    bExecute : BOOL;
    tTimeout : TIME := T#2S;
END_VAR
VAR_OUTPUT
    bBusy : BOOL;
    bDone : BOOL;
    bError : BOOL;
    nErrId : UDINT;
    nStatus : DINT;
    bAuthed : BOOL;
    sValue : STRING[127];        // query: current input number
END_VAR
VAR
    pjl : FB_PJLink;
END_VAR
    pjl.sHost := sHost;
    pjl.nPort := nPort;
    pjl.nCls := 1;
    pjl.sCmd := 'INPT';
    IF nMode = 1 THEN
        pjl.sParam := '?';
    ELSE
        pjl.sParam := sInput;
    END_IF;
    pjl.sPassword := sPassword;
    pjl.tTimeout := tTimeout;
    pjl.bExecute := bExecute;
    pjl();
    bBusy := pjl.bBusy;
    bDone := pjl.bDone;
    bError := pjl.bError;
    nErrId := pjl.nErrId;
    nStatus := pjl.nStatus;
    bAuthed := pjl.bAuthed;
    sValue := pjl.sValue;
END_FUNCTION_BLOCK

// AV mute on/off/query — TwinCAT SetMute/QueryMute methods.
// PJLink AVMT: 30=mute off (open), 31=mute on (closed);
// query returns 11/21/30/31.
FUNCTION_BLOCK FB_PJLink_Mute
VAR_INPUT
    sHost : STRING[15];
    nPort : UDINT := 4352;
    sPassword : STRING[32] := '';
    nMode : UDINT;               // 0=mute on 1=mute off 2=query
    bExecute : BOOL;
    tTimeout : TIME := T#2S;
END_VAR
VAR_OUTPUT
    bBusy : BOOL;
    bDone : BOOL;
    bError : BOOL;
    nErrId : UDINT;
    nStatus : DINT;
    bAuthed : BOOL;
    sValue : STRING[127];        // query: "11"/"21"/"30"/"31"
END_VAR
VAR
    pjl : FB_PJLink;
END_VAR
    pjl.sHost := sHost;
    pjl.nPort := nPort;
    pjl.nCls := 1;
    pjl.sCmd := 'AVMT';
    IF nMode = 2 THEN
        pjl.sParam := '?';
    ELSIF nMode = 0 THEN
        pjl.sParam := '31';
    ELSE
        pjl.sParam := '30';
    END_IF;
    pjl.sPassword := sPassword;
    pjl.tTimeout := tTimeout;
    pjl.bExecute := bExecute;
    pjl();
    bBusy := pjl.bBusy;
    bDone := pjl.bDone;
    bError := pjl.bError;
    nErrId := pjl.nErrId;
    nStatus := pjl.nStatus;
    bAuthed := pjl.bAuthed;
    sValue := pjl.sValue;
END_FUNCTION_BLOCK

(* ---- tc3_plctest.st ---- *)
// Tc3_PlcTestFramework (TF1140) -> PLC-side test framework.
// Beckhoff's library exposes a METHOD-based assertion API on
// FB_TestCaseBase/FB_TestPrepBase plus a test client that drives
// the run.  This port keeps the assertion/step semantics and
// replaces the METHOD calls with edge-triggered command inputs
// (this compiler has no METHOD support):
//   FB_TestCase   nAssertCmd 1=Assert 2=AssertEqual
//                 3=AssertAbsEqual 4=AssertRelEqual
//                 5=AssertStrictLarger
//                 nCmd 1=IncStep 2=GoToStep 3=IncStepIf 4=Cleanup
//                 5=Reset
//   FB_TestSuite  nCmd 1=AddResult 2=Reset
// Documented differences:
//   - No test client / no .tcuitest files: results are PLC values
//     (counters + bSucceeded) that the host or a CI script reads
//     from the process image.
//   - Assertions are counted, not reported with stack traces;
//     nFailures is the failure count and bSucceeded the verdict.
//   - AssertMsg carries no message text (documented reduction).

FUNCTION_BLOCK FB_TestCase
VAR_INPUT
    // assertion request
    nAssertCmd : UDINT;         // see header
    bAssertCond : BOOL;         // Assert / AssertMsg
    fActual : LREAL;
    fExpected : LREAL;
    fTolerance : LREAL;         // abs tolerance / rel fraction
    // step control
    nCmd : UDINT;
    nStepArg : UDINT;
    bStepCond : BOOL;           // IncStepIf
END_VAR
VAR_OUTPUT
    nAssertions : UDINT;
    nFailures : UDINT;
    nStep : UDINT;
    bSucceeded : BOOL;
    bDone : BOOL;
    bError : BOOL;
    nErrId : UDINT;
END_VAR
VAR
    prevAssert : UDINT;
    prevCmd : UDINT;
    fDiff : LREAL;
    fRel : LREAL;
    ok : BOOL;
END_VAR
    bDone := FALSE; bError := FALSE; nErrId := 0;

    // ---- assertions ----
    IF nAssertCmd <> 0 AND prevAssert = 0 THEN
        ok := FALSE;
        IF nAssertCmd = 1 THEN
            ok := bAssertCond;
        ELSIF nAssertCmd = 2 THEN
            ok := fActual = fExpected;
        ELSIF nAssertCmd = 3 THEN
            fDiff := fActual - fExpected;
            IF fDiff < 0.0 THEN fDiff := -fDiff; END_IF;
            ok := fDiff <= fTolerance;
        ELSIF nAssertCmd = 4 THEN
            fRel := 0.0;
            IF fExpected <> 0.0 THEN
                fRel := (fActual - fExpected) / fExpected;
                IF fRel < 0.0 THEN fRel := -fRel; END_IF;
            END_IF;
            ok := fRel <= fTolerance;
        ELSIF nAssertCmd = 5 THEN
            ok := fActual > fExpected;
        END_IF;
        nAssertions := nAssertions + 1;
        IF NOT ok THEN nFailures := nFailures + 1; END_IF;
        bDone := TRUE;
    END_IF;
    prevAssert := nAssertCmd;

    // ---- step control ----
    IF nCmd <> 0 AND prevCmd = 0 THEN
        IF nCmd = 1 THEN
            nStep := nStep + 1;
            bDone := TRUE;
        ELSIF nCmd = 2 THEN
            nStep := nStepArg;
            bDone := TRUE;
        ELSIF nCmd = 3 THEN
            IF bStepCond THEN nStep := nStep + 1; END_IF;
            bDone := TRUE;
        ELSIF nCmd = 4 THEN
            bDone := TRUE;          // Cleanup: nothing owned here
        ELSIF nCmd = 5 THEN
            nStep := 0; nAssertions := 0; nFailures := 0;
            bDone := TRUE;
        ELSE
            bError := TRUE; nErrId := 1;
        END_IF;
    END_IF;
    prevCmd := nCmd;

    bSucceeded := nFailures = 0;
END_FUNCTION_BLOCK

// ---- FB_TestPrepBase: same surface, used for fixtures ----
// The upstream Prep block differs only in the run phase; here it is
// the same implementation with a distinct type so suites can tell
// preparation assertions from test assertions.
FUNCTION_BLOCK FB_TestPrepBase
VAR_INPUT
    nAssertCmd : UDINT;
    bAssertCond : BOOL;
    fActual : LREAL;
    fExpected : LREAL;
    fTolerance : LREAL;
    nCmd : UDINT;
    nStepArg : UDINT;
    bStepCond : BOOL;
END_VAR
VAR_OUTPUT
    nAssertions : UDINT;
    nFailures : UDINT;
    nStep : UDINT;
    bSucceeded : BOOL;
    bDone : BOOL;
    bError : BOOL;
    nErrId : UDINT;
END_VAR
VAR
    tc : FB_TestCase;
END_VAR
    tc.nAssertCmd := nAssertCmd;
    tc.bAssertCond := bAssertCond;
    tc.fActual := fActual;
    tc.fExpected := fExpected;
    tc.fTolerance := fTolerance;
    tc.nCmd := nCmd;
    tc.nStepArg := nStepArg;
    tc.bStepCond := bStepCond;
    tc();
    nAssertions := tc.nAssertions;
    nFailures := tc.nFailures;
    nStep := tc.nStep;
    bSucceeded := tc.bSucceeded;
    bDone := tc.bDone;
    bError := tc.bError;
    nErrId := tc.nErrId;
END_FUNCTION_BLOCK

// ---- FB_TestCaseBasePrep: prep-phase variant of the case ----
FUNCTION_BLOCK FB_TestCaseBasePrep
VAR_INPUT
    nAssertCmd : UDINT;
    bAssertCond : BOOL;
    fActual : LREAL;
    fExpected : LREAL;
    fTolerance : LREAL;
    nCmd : UDINT;
    nStepArg : UDINT;
    bStepCond : BOOL;
END_VAR
VAR_OUTPUT
    nAssertions : UDINT;
    nFailures : UDINT;
    nStep : UDINT;
    bSucceeded : BOOL;
    bDone : BOOL;
    bError : BOOL;
    nErrId : UDINT;
END_VAR
VAR
    tc : FB_TestCase;
END_VAR
    tc.nAssertCmd := nAssertCmd;
    tc.bAssertCond := bAssertCond;
    tc.fActual := fActual;
    tc.fExpected := fExpected;
    tc.fTolerance := fTolerance;
    tc.nCmd := nCmd;
    tc.nStepArg := nStepArg;
    tc.bStepCond := bStepCond;
    tc();
    nAssertions := tc.nAssertions;
    nFailures := tc.nFailures;
    nStep := tc.nStep;
    bSucceeded := tc.bSucceeded;
    bDone := tc.bDone;
    bError := tc.bError;
    nErrId := tc.nErrId;
END_FUNCTION_BLOCK

// ---- FB_TestSuite: aggregate case results ----
FUNCTION_BLOCK FB_TestSuite
VAR_INPUT
    nCmd : UDINT;               // 1=AddResult 2=Reset
    bCasePassed : BOOL;
END_VAR
VAR_OUTPUT
    nTests : UDINT;
    nPassed : UDINT;
    nFailed : UDINT;
    bAllPassed : BOOL;
    bDone : BOOL;
END_VAR
VAR
    prev : UDINT;
END_VAR
    bDone := FALSE;
    IF nCmd <> 0 AND prev = 0 THEN
        IF nCmd = 1 THEN
            nTests := nTests + 1;
            IF bCasePassed THEN
                nPassed := nPassed + 1;
            ELSE
                nFailed := nFailed + 1;
            END_IF;
            bDone := TRUE;
        ELSIF nCmd = 2 THEN
            nTests := 0; nPassed := 0; nFailed := 0;
            bDone := TRUE;
        END_IF;
    END_IF;
    prev := nCmd;
    bAllPassed := nFailed = 0 AND nTests > 0;
END_FUNCTION_BLOCK

(* ---- tc3_robotics.st ---- *)
// tc3_robotics.st — Tc3_mxAutomation (TF5120, KUKA.PLC mxA) and
// Tc3_uniValPlc (TF5130, Stäubli uniVAL plc) surfaces.  Both are
// licensed Beckhoff robotics engines talking to proprietary robot
// controllers; TetherPLC ships neither engine nor license, so
// these blocks are honest license/engine-absent stubs: commands
// are validated (bad inputs fail immediately), Busy runs a
// bounded handshake, then Error with a documented ErrorId — no
// robot state, motion, or I/O result is ever faked.
//
// Differences (docs/plc/compat/README.md):
//   - mxAutomation's FB_KRC_Group / FB_KRC_Move* family and
//     uniVAL's FB_Val3 group/command family are unified here as
//     FB_RobotGroup (connect/poll) and FB_RobotCommand
//     (PTP/LIN/CIRC dispatch) — the proprietary protocol surfaces
//     (mxA telegram, uniVAL CS8/CS9) have no backend.
//   - ErrorId: 0 none, 1 engine/license-unavailable,
//     2 bad-address, 3 bad-move, 4 aborted, 5 not-connected.

// ---- FB_RobotGroup: robot-controller group connection ----
// Covers FB_KRC_Group.Open/Disconnect and FB_Val3 group attach.
FUNCTION_BLOCK FB_RobotGroup
VAR_INPUT
    Connect : BOOL;             // rising edge opens the session
    Disconnect : BOOL;
    Controller : STRING;        // controller address/endpoint
    RobotCount : UDINT;         // robots in the group (>=1)
END_VAR
VAR_OUTPUT
    Connected : BOOL;
    Busy : BOOL;
    Error : BOOL;
    ErrorId : UDINT;
END_VAR
VAR
    phase : INT;
    tmo : UDINT;
END_VAR
    IF phase = 0 THEN
        Busy := FALSE;
        IF Connect THEN
            Busy := TRUE;
            Error := FALSE;
            ErrorId := 0;
            Connected := FALSE;
            tmo := 0;
            IF Controller = '' OR RobotCount = 0 THEN
                Error := TRUE;
                ErrorId := 2;        // bad-address
                Busy := FALSE;
                phase := 2;
            ELSE
                phase := 1;
            END_IF;
        END_IF;
    ELSIF phase = 1 THEN
        tmo := tmo + 1;
        IF tmo >= 4 THEN
            Busy := FALSE;
            Error := TRUE;
            ErrorId := 1;            // license/engine unavailable
            phase := 2;
        END_IF;
    ELSE
        Busy := FALSE;
        IF NOT Connect THEN
            phase := 0;
        END_IF;
    END_IF;
    IF Disconnect THEN
        Connected := FALSE;
        Busy := FALSE;
        phase := 0;
    END_IF;
END_FUNCTION_BLOCK

// ---- FB_RobotCommand: PTP/LIN/CIRC motion dispatch ----
// Covers the FB_KRC_Move*/FB_Val3Move* async-command spine.
FUNCTION_BLOCK FB_RobotCommand
VAR_INPUT
    Execute : BOOL;
    Abort : BOOL;
    GroupConnected : BOOL;      // from FB_RobotGroup.Connected
    MoveType : UDINT;           // 1 PTP, 2 LIN, 3 CIRC
    X : LREAL; Y : LREAL; Z : LREAL;
    Velocity : LREAL;           // mm/s or % override (>0)
END_VAR
VAR_OUTPUT
    Busy : BOOL;
    Active : BOOL;
    Done : BOOL;
    CommandAborted : BOOL;
    Error : BOOL;
    ErrorId : UDINT;
    ReachedTarget : BOOL;        // never TRUE without an engine
END_VAR
VAR
    phase : INT;
    tmo : UDINT;
END_VAR
    Done := FALSE;
    Active := FALSE;
    CommandAborted := FALSE;
    ReachedTarget := FALSE;
    IF phase = 0 THEN
        Busy := FALSE;
        IF Execute THEN
            Busy := TRUE;
            Active := TRUE;
            Error := FALSE;
            ErrorId := 0;
            tmo := 0;
            IF NOT GroupConnected THEN
                Error := TRUE;
                ErrorId := 5;        // not-connected
                Active := FALSE;
                Busy := FALSE;
                phase := 2;
            ELSIF MoveType = 0 OR MoveType > 3 OR Velocity <= 0.0 THEN
                Error := TRUE;
                ErrorId := 3;        // bad-move
                Active := FALSE;
                Busy := FALSE;
                phase := 2;
            ELSE
                phase := 1;
            END_IF;
        END_IF;
    ELSIF phase = 1 THEN
        tmo := tmo + 1;
        IF tmo >= 4 THEN
            Busy := FALSE;
            Active := FALSE;
            Error := TRUE;
            ErrorId := 1;            // license/engine unavailable
            phase := 2;
        END_IF;
    ELSE
        Busy := FALSE;
        IF NOT Execute THEN
            phase := 0;
        END_IF;
    END_IF;
    IF Abort AND phase = 1 THEN
        Busy := FALSE;
        Active := FALSE;
        CommandAborted := TRUE;
        Error := TRUE;
        ErrorId := 4;
        phase := 2;
    END_IF;
    Done := (phase = 2);
END_FUNCTION_BLOCK

(* ---- tc3_rtmon.st ---- *)
// Tc3_RealtimeMonitoring compatibility (TwinCAT 3 PLC Library
// Tc3_RealtimeMonitoring). Beckhoff-shaped wrappers over the builtin
// FB_RtMon, which drives the host "tplc-rtmon" service: a bounded
// ring of timestamped marks (steady-clock ns; sim time under
// --sim), appended from the scan path.
//
// Differences from TwinCAT, documented in docs/plc/compat/README.md:
//   - TwinCAT exposes methods on the FBs (fb.LogMark(...)); this
//     dialect has no METHOD, so each method is a separate
//     FUNCTION_BLOCK gated by bExecute: one rising edge = one mark.
//   - nContextId default TwinCAT_SystemInfoVarList._AppInfo.AdsPort
//     is unavailable; pass the context explicitly.
//   - bLogCallingTask / TcMarkOption.RefToCaller only records the
//     flag bit in the stored markctrl; no task reference is resolved.
//   - FB_RTMon_LogTrigger stores a plain mark; the realtime-monitor
//     server-side recording trigger is not modeled.
//   - hrErrorCode carries 0 or a negative service code, not a real
//     COM HRESULT.
//   - TcMarkOption has no VAR_GLOBAL CONSTANT in this dialect; the
//     UDINT masks are documented inline at each call site:
//       Start            16#E0000000   Stop             16#C0000000
//       SequenceStart    16#A0000000   SequenceStop     16#80000000
//       IntervalStart    16#60000000   IntervalStop     16#40000000
//       RefToCaller      16#08000000   (OR with a type)
//   - ST_RTMon_MarkDef cannot cross the --lib boundary (types are
//     file-scoped in this dialect), so LogMarkEx takes the three
//     MarkDef fields (nContextId/nGroupId/nEventId) flattened.
// Sources: docs/plc/plan/21-twincat-libraries.md §7 (TE1010).

// ---- FB_RTMon_LogMarkBase family (explicit context + markctrl) ----

FUNCTION_BLOCK FB_RTMon_LogMarkBase
VAR_INPUT
    bExecute : BOOL;
    nContextId : UINT;
    nGroupId : UINT;
    nEventId : UINT;
    nMarkCtrl : UDINT;
END_VAR
VAR_OUTPUT
    bBusy : BOOL;
    bDone : BOOL;
    bError : BOOL;
    hrErrorCode : DINT;
END_VAR
VAR
    rtmon : FB_RtMon;
END_VAR
    rtmon.OP := 1;
    rtmon.CONTEXT := nContextId;
    rtmon.GROUP := nGroupId;
    rtmon.EVENT := nEventId;
    rtmon.MARKCTRL := nMarkCtrl;
    rtmon.EXEC := bExecute;
    rtmon();
    bBusy := rtmon.BUSY;
    bDone := rtmon.DONE;
    bError := rtmon.ERRID <> 0;
    hrErrorCode := rtmon.RESULT - UDINT_TO_DINT(rtmon.ERRID);
END_FUNCTION_BLOCK

// FB_RTMon_LogMarkBase.LogMarkEx — stMark flattened to its three
// UINT fields (see header note on ST_RTMon_MarkDef).
FUNCTION_BLOCK FB_RTMon_LogMarkBaseEx
VAR_INPUT
    bExecute : BOOL;
    nContextId : UINT;
    nGroupId : UINT;
    nEventId : UINT;
    nMarkCtrl : UDINT;
END_VAR
VAR_OUTPUT
    bBusy : BOOL;
    bDone : BOOL;
    bError : BOOL;
    hrErrorCode : DINT;
END_VAR
VAR
    rtmon : FB_RtMon;
END_VAR
    rtmon.OP := 1;
    rtmon.CONTEXT := nContextId;
    rtmon.GROUP := nGroupId;
    rtmon.EVENT := nEventId;
    rtmon.MARKCTRL := nMarkCtrl;
    rtmon.EXEC := bExecute;
    rtmon();
    bBusy := rtmon.BUSY;
    bDone := rtmon.DONE;
    bError := rtmon.ERRID <> 0;
    hrErrorCode := rtmon.RESULT - UDINT_TO_DINT(rtmon.ERRID);
END_FUNCTION_BLOCK

// ---- FB_RTMon_LogMark family (context on the call, fixed type) ----
// Each FB embeds the markctrl for its TwinCAT method; bLogCallingTask
// ORs in TcMarkOption.RefToCaller (16#08000000).

FUNCTION_BLOCK FB_RTMon_LogMark
VAR_INPUT
    bExecute : BOOL;
    nContextId : UINT;
    bLogCallingTask : BOOL := TRUE;
    nGroupId : UINT;
    nEventId : UINT;
END_VAR
VAR_OUTPUT
    bBusy : BOOL;
    bDone : BOOL;
    bError : BOOL;
    hrErrorCode : DINT;
END_VAR
VAR
    rtmon : FB_RtMon;
    mctrl : UDINT;
END_VAR
    mctrl := 16#00000000;
    IF bLogCallingTask THEN
        mctrl := mctrl + 16#08000000;
    END_IF;
    rtmon.OP := 1;
    rtmon.CONTEXT := nContextId;
    rtmon.GROUP := nGroupId;
    rtmon.EVENT := nEventId;
    rtmon.MARKCTRL := mctrl;
    rtmon.EXEC := bExecute;
    rtmon();
    bBusy := rtmon.BUSY;
    bDone := rtmon.DONE;
    bError := rtmon.ERRID <> 0;
    hrErrorCode := rtmon.RESULT - UDINT_TO_DINT(rtmon.ERRID);
END_FUNCTION_BLOCK

FUNCTION_BLOCK FB_RTMon_LogIntervalStart
VAR_INPUT
    bExecute : BOOL;
    nContextId : UINT;
    bLogCallingTask : BOOL := TRUE;
    nGroupId : UINT;
    nEventId : UINT;
END_VAR
VAR_OUTPUT
    bBusy : BOOL;
    bDone : BOOL;
    bError : BOOL;
    hrErrorCode : DINT;
END_VAR
VAR
    rtmon : FB_RtMon;
    mctrl : UDINT;
END_VAR
    mctrl := 16#60000000;
    IF bLogCallingTask THEN
        mctrl := mctrl + 16#08000000;
    END_IF;
    rtmon.OP := 1;
    rtmon.CONTEXT := nContextId;
    rtmon.GROUP := nGroupId;
    rtmon.EVENT := nEventId;
    rtmon.MARKCTRL := mctrl;
    rtmon.EXEC := bExecute;
    rtmon();
    bBusy := rtmon.BUSY;
    bDone := rtmon.DONE;
    bError := rtmon.ERRID <> 0;
    hrErrorCode := rtmon.RESULT - UDINT_TO_DINT(rtmon.ERRID);
END_FUNCTION_BLOCK

FUNCTION_BLOCK FB_RTMon_LogIntervalStop
VAR_INPUT
    bExecute : BOOL;
    nContextId : UINT;
    bLogCallingTask : BOOL := TRUE;
    nGroupId : UINT;
    nEventId : UINT;
END_VAR
VAR_OUTPUT
    bBusy : BOOL;
    bDone : BOOL;
    bError : BOOL;
    hrErrorCode : DINT;
END_VAR
VAR
    rtmon : FB_RtMon;
    mctrl : UDINT;
END_VAR
    mctrl := 16#40000000;
    IF bLogCallingTask THEN
        mctrl := mctrl + 16#08000000;
    END_IF;
    rtmon.OP := 1;
    rtmon.CONTEXT := nContextId;
    rtmon.GROUP := nGroupId;
    rtmon.EVENT := nEventId;
    rtmon.MARKCTRL := mctrl;
    rtmon.EXEC := bExecute;
    rtmon();
    bBusy := rtmon.BUSY;
    bDone := rtmon.DONE;
    bError := rtmon.ERRID <> 0;
    hrErrorCode := rtmon.RESULT - UDINT_TO_DINT(rtmon.ERRID);
END_FUNCTION_BLOCK

FUNCTION_BLOCK FB_RTMon_LogSequenceStart
VAR_INPUT
    bExecute : BOOL;
    nContextId : UINT;
    bLogCallingTask : BOOL := TRUE;
    nGroupId : UINT;
    nEventId : UINT;
END_VAR
VAR_OUTPUT
    bBusy : BOOL;
    bDone : BOOL;
    bError : BOOL;
    hrErrorCode : DINT;
END_VAR
VAR
    rtmon : FB_RtMon;
    mctrl : UDINT;
END_VAR
    mctrl := 16#A0000000;
    IF bLogCallingTask THEN
        mctrl := mctrl + 16#08000000;
    END_IF;
    rtmon.OP := 1;
    rtmon.CONTEXT := nContextId;
    rtmon.GROUP := nGroupId;
    rtmon.EVENT := nEventId;
    rtmon.MARKCTRL := mctrl;
    rtmon.EXEC := bExecute;
    rtmon();
    bBusy := rtmon.BUSY;
    bDone := rtmon.DONE;
    bError := rtmon.ERRID <> 0;
    hrErrorCode := rtmon.RESULT - UDINT_TO_DINT(rtmon.ERRID);
END_FUNCTION_BLOCK

FUNCTION_BLOCK FB_RTMon_LogSequenceStop
VAR_INPUT
    bExecute : BOOL;
    nContextId : UINT;
    bLogCallingTask : BOOL := TRUE;
    nGroupId : UINT;
    nEventId : UINT;
END_VAR
VAR_OUTPUT
    bBusy : BOOL;
    bDone : BOOL;
    bError : BOOL;
    hrErrorCode : DINT;
END_VAR
VAR
    rtmon : FB_RtMon;
    mctrl : UDINT;
END_VAR
    mctrl := 16#80000000;
    IF bLogCallingTask THEN
        mctrl := mctrl + 16#08000000;
    END_IF;
    rtmon.OP := 1;
    rtmon.CONTEXT := nContextId;
    rtmon.GROUP := nGroupId;
    rtmon.EVENT := nEventId;
    rtmon.MARKCTRL := mctrl;
    rtmon.EXEC := bExecute;
    rtmon();
    bBusy := rtmon.BUSY;
    bDone := rtmon.DONE;
    bError := rtmon.ERRID <> 0;
    hrErrorCode := rtmon.RESULT - UDINT_TO_DINT(rtmon.ERRID);
END_FUNCTION_BLOCK

FUNCTION_BLOCK FB_RTMon_LogStart
VAR_INPUT
    bExecute : BOOL;
    nContextId : UINT;
    bLogCallingTask : BOOL := TRUE;
    nGroupId : UINT;
    nEventId : UINT;
END_VAR
VAR_OUTPUT
    bBusy : BOOL;
    bDone : BOOL;
    bError : BOOL;
    hrErrorCode : DINT;
END_VAR
VAR
    rtmon : FB_RtMon;
    mctrl : UDINT;
END_VAR
    mctrl := 16#E0000000;
    IF bLogCallingTask THEN
        mctrl := mctrl + 16#08000000;
    END_IF;
    rtmon.OP := 1;
    rtmon.CONTEXT := nContextId;
    rtmon.GROUP := nGroupId;
    rtmon.EVENT := nEventId;
    rtmon.MARKCTRL := mctrl;
    rtmon.EXEC := bExecute;
    rtmon();
    bBusy := rtmon.BUSY;
    bDone := rtmon.DONE;
    bError := rtmon.ERRID <> 0;
    hrErrorCode := rtmon.RESULT - UDINT_TO_DINT(rtmon.ERRID);
END_FUNCTION_BLOCK

FUNCTION_BLOCK FB_RTMon_LogStop
VAR_INPUT
    bExecute : BOOL;
    nContextId : UINT;
    bLogCallingTask : BOOL := TRUE;
    nGroupId : UINT;
    nEventId : UINT;
END_VAR
VAR_OUTPUT
    bBusy : BOOL;
    bDone : BOOL;
    bError : BOOL;
    hrErrorCode : DINT;
END_VAR
VAR
    rtmon : FB_RtMon;
    mctrl : UDINT;
END_VAR
    mctrl := 16#C0000000;
    IF bLogCallingTask THEN
        mctrl := mctrl + 16#08000000;
    END_IF;
    rtmon.OP := 1;
    rtmon.CONTEXT := nContextId;
    rtmon.GROUP := nGroupId;
    rtmon.EVENT := nEventId;
    rtmon.MARKCTRL := mctrl;
    rtmon.EXEC := bExecute;
    rtmon();
    bBusy := rtmon.BUSY;
    bDone := rtmon.DONE;
    bError := rtmon.ERRID <> 0;
    hrErrorCode := rtmon.RESULT - UDINT_TO_DINT(rtmon.ERRID);
END_FUNCTION_BLOCK

FUNCTION_BLOCK FB_RTMon_LogTrigger
VAR_INPUT
    bExecute : BOOL;
    nContextId : UINT;
    bLogCallingTask : BOOL := TRUE;
    nGroupId : UINT;
    nEventId : UINT;
END_VAR
VAR_OUTPUT
    bBusy : BOOL;
    bDone : BOOL;
    bError : BOOL;
    hrErrorCode : DINT;
END_VAR
VAR
    rtmon : FB_RtMon;
    mctrl : UDINT;
END_VAR
    // TwinCAT trigger marks arm server-side recording; with no
    // trigger bit defined we store a plain mark (markctrl 0)
    mctrl := 16#00000000;
    IF bLogCallingTask THEN
        mctrl := mctrl + 16#08000000;
    END_IF;
    rtmon.OP := 1;
    rtmon.CONTEXT := nContextId;
    rtmon.GROUP := nGroupId;
    rtmon.EVENT := nEventId;
    rtmon.MARKCTRL := mctrl;
    rtmon.EXEC := bExecute;
    rtmon();
    bBusy := rtmon.BUSY;
    bDone := rtmon.DONE;
    bError := rtmon.ERRID <> 0;
    hrErrorCode := rtmon.RESULT - UDINT_TO_DINT(rtmon.ERRID);
END_FUNCTION_BLOCK

(* ---- tc3_s7comm.st ---- *)
// Tc3_S7Comm + Tc2_S5S7Com -> Siemens S7comm client wrappers.
// TwinCAT's FB_S7CommConnection owns an AMS-routed session with
// I_S7CommRequest objects, PVOID buffers and HRESULT returns;
// Tc2_S5S7Com's FB_NLink* blocks map fetch/write requests onto
// T_HNLINK handles. TetherPLC adapts both to the poll-driven
// service model used by the other compat libraries: FB_S7Conn
// holds the persistent RFC1006/COTP session, FB_S7Io runs one
// Read Var / Write Var transaction per EXEC edge.
// Differences from the TwinCAT FBs, documented in
// docs/plc/compat/README.md:
//   - No AMS NetID routing, no PVOID/HRESULT/interface request
//     objects, no cyclic request queues (AddRequest* variants).
//     Requests are explicit poll-model FBs; one outstanding
//     transaction per connection.
//   - IPv4 dotted-quad hosts only, no DNS.
//   - nArea is the raw S7-Any area code: 16#81=PE(I), 16#82=PA(Q),
//     16#83=MK(M), 16#84=DB, 16#1C=CT, 16#1D=TM.
//   - nStatus: conn 0=pending 1=ready 2=error; io 0=pending
//     1=ok 2=timeout 3=error 4=badresp 5=s7err. nErrId carries
//     the transport errno or S7 error word; nItemRc the response
//     item return code (16#FF ok).
//   - Bit reads return one byte in pData[0] with the bit value
//     right-justified (bit 0); bit writes take pData[0]&1.
// Sources: docs/plc/plan/21-twincat-libraries.md (Tc2_S5S7Com,
// Tc3_S7Comm).

// Open/poll/close a persistent S7 connection — covers
// FB_S7CommConnection and the FB_NLinkOpen/FB_NLinkClose pair.
FUNCTION_BLOCK FB_S7_Connect
VAR_INPUT
    sHost : STRING[15];          // dotted-quad PLC IPv4
    nPort : UDINT := 0;          // 0 = 102
    nRack : UDINT := 0;          // 0..15
    nSlot : UDINT := 2;          // 0..31
    bExecute : BOOL;             // rising edge = (re)connect
    bClose : BOOL;               // rising edge = disconnect
    tTimeout : TIME := T#5S;
END_VAR
VAR_OUTPUT
    nConnHandle : UDINT;         // 0 = no live session
    bBusy : BOOL;
    bDone : BOOL;
    bError : BOOL;
    nStatus : DINT;              // 0=pending 1=ready 2=error
    nErrId : UDINT;
END_VAR
VAR
    conn : FB_S7Conn;
END_VAR
    conn.HOST := sHost;
    conn.PORT := nPort;
    conn.RACK := nRack;
    conn.SLOT := nSlot;
    conn.TIMEOUT := tTimeout;
    conn.CLOSE := bClose;
    conn.EXEC := bExecute;
    conn();
    nConnHandle := conn.CONN_HANDLE;
    bBusy := conn.BUSY;
    bDone := conn.DONE;
    nStatus := conn.STATUS;
    nErrId := conn.ERRID;
    bError := (conn.ERRID <> 0) OR (conn.STATUS = 2);
END_FUNCTION_BLOCK

// Read bytes — covers FB_S7CommCyclicRequest/AddReadVar/
// AddReadByteArray and FB_NLinkFetch.
FUNCTION_BLOCK FB_S7_Read
VAR_INPUT
    nConnHandle : UDINT;         // from FB_S7_Connect
    nArea : UDINT;               // S7-Any area code
    nDb : UDINT := 0;            // DB number (DB area only)
    nByteOff : UDINT;            // byte offset (24-bit)
    nLen : UDINT;                // bytes, 1..240
    bExecute : BOOL;
    tTimeout : TIME := T#2S;
END_VAR
VAR_OUTPUT
    bBusy : BOOL;
    bDone : BOOL;
    bError : BOOL;
    nErrId : UDINT;
    nStatus : DINT;              // 0=pending 1=ok 2=timeout 3=err
                                  // 4=badresp 5=s7err
    nItemRc : UDINT;             // response item return code
    nDataLen : UDINT;            // valid bytes in pData
    pData : ARRAY[0..239] OF BYTE;
END_VAR
VAR
    io : FB_S7Io;
    i : UDINT;
END_VAR
    io.CONN_HANDLE := nConnHandle;
    io.MODE := 0;
    io.AREA := nArea;
    io.DB := nDb;
    io.BYTE_OFF := nByteOff;
    io.BIT_ACCESS := FALSE;
    io.BIT_NO := 0;
    io.LEN := nLen;
    io.TIMEOUT := tTimeout;
    io.EXEC := bExecute;
    io();
    bBusy := io.BUSY;
    bDone := io.DONE;
    nStatus := io.STATUS;
    nErrId := io.ERRID;
    nItemRc := io.ITEM_RC;
    nDataLen := io.DATA_LEN;
    IF io.DONE THEN
        i := 0;
        WHILE i < io.DATA_LEN AND i < 240 DO
            pData[i] := io.R_DATA[i];
            i := i + 1;
        END_WHILE;
    END_IF;
    bError := (io.ERRID <> 0) OR (io.STATUS >= 2);
END_FUNCTION_BLOCK

// Write bytes — covers AddWriteVar/AddWriteByteArray and
// FB_NLinkWrite.
FUNCTION_BLOCK FB_S7_Write
VAR_INPUT
    nConnHandle : UDINT;
    nArea : UDINT;
    nDb : UDINT := 0;
    nByteOff : UDINT;
    nLen : UDINT;                // bytes, 1..240
    pData : ARRAY[0..239] OF BYTE;
    bExecute : BOOL;
    tTimeout : TIME := T#2S;
END_VAR
VAR_OUTPUT
    bBusy : BOOL;
    bDone : BOOL;
    bError : BOOL;
    nErrId : UDINT;
    nStatus : DINT;
    nItemRc : UDINT;
END_VAR
VAR
    io : FB_S7Io;
    i : UDINT;
END_VAR
    io.CONN_HANDLE := nConnHandle;
    io.MODE := 1;
    io.AREA := nArea;
    io.DB := nDb;
    io.BYTE_OFF := nByteOff;
    io.BIT_ACCESS := FALSE;
    io.BIT_NO := 0;
    io.LEN := nLen;
    io.TIMEOUT := tTimeout;
    i := 0;
    WHILE i < nLen AND i < 240 DO
        io.DATA[i] := pData[i];
        i := i + 1;
    END_WHILE;
    io.EXEC := bExecute;
    io();
    bBusy := io.BUSY;
    bDone := io.DONE;
    nStatus := io.STATUS;
    nErrId := io.ERRID;
    nItemRc := io.ITEM_RC;
    bError := (io.ERRID <> 0) OR (io.STATUS >= 2);
END_FUNCTION_BLOCK

// Read one bit — covers AddReadBit. nBitNo 0..7 selects the bit
// inside nByteOff; pData[0] bit 0 holds the value when done.
FUNCTION_BLOCK FB_S7_ReadBit
VAR_INPUT
    nConnHandle : UDINT;
    nArea : UDINT;
    nDb : UDINT := 0;
    nByteOff : UDINT;
    nBitNo : UDINT;              // 0..7
    bExecute : BOOL;
    tTimeout : TIME := T#2S;
END_VAR
VAR_OUTPUT
    bBusy : BOOL;
    bDone : BOOL;
    bError : BOOL;
    nErrId : UDINT;
    nStatus : DINT;
    nItemRc : UDINT;
    nBitValue : UDINT;           // 0 or 1
END_VAR
VAR
    io : FB_S7Io;
END_VAR
    io.CONN_HANDLE := nConnHandle;
    io.MODE := 0;
    io.AREA := nArea;
    io.DB := nDb;
    io.BYTE_OFF := nByteOff;
    io.BIT_ACCESS := TRUE;
    io.BIT_NO := nBitNo;
    io.LEN := 1;
    io.TIMEOUT := tTimeout;
    io.EXEC := bExecute;
    io();
    bBusy := io.BUSY;
    bDone := io.DONE;
    nStatus := io.STATUS;
    nErrId := io.ERRID;
    nItemRc := io.ITEM_RC;
    IF io.DONE AND io.STATUS = 1 THEN
        nBitValue := BYTE_TO_UDINT(io.R_DATA[0]) AND 16#01;
    ELSE
        nBitValue := 0;
    END_IF;
    bError := (io.ERRID <> 0) OR (io.STATUS >= 2);
END_FUNCTION_BLOCK

// Write one bit — covers the AddWrite* bit variants.
// nBitValue 0 clears, nonzero sets.
FUNCTION_BLOCK FB_S7_WriteBit
VAR_INPUT
    nConnHandle : UDINT;
    nArea : UDINT;
    nDb : UDINT := 0;
    nByteOff : UDINT;
    nBitNo : UDINT;              // 0..7
    nBitValue : UDINT;           // 0 or 1
    bExecute : BOOL;
    tTimeout : TIME := T#2S;
END_VAR
VAR_OUTPUT
    bBusy : BOOL;
    bDone : BOOL;
    bError : BOOL;
    nErrId : UDINT;
    nStatus : DINT;
    nItemRc : UDINT;
END_VAR
VAR
    io : FB_S7Io;
END_VAR
    io.CONN_HANDLE := nConnHandle;
    io.MODE := 1;
    io.AREA := nArea;
    io.DB := nDb;
    io.BYTE_OFF := nByteOff;
    io.BIT_ACCESS := TRUE;
    io.BIT_NO := nBitNo;
    io.LEN := 1;
    io.TIMEOUT := tTimeout;
    io.DATA[0] := UDINT_TO_BYTE(nBitValue AND 16#01);
    io.EXEC := bExecute;
    io();
    bBusy := io.BUSY;
    bDone := io.DONE;
    nStatus := io.STATUS;
    nErrId := io.ERRID;
    nItemRc := io.ITEM_RC;
    bError := (io.ERRID <> 0) OR (io.STATUS >= 2);
END_FUNCTION_BLOCK

(* ---- tc3_sacn.st ---- *)
// Tc3_sACN compatibility (TwinCAT 3 PLC Library Tc3_sACN, ANSI
// E1.31 streaming ACN). Beckhoff-shaped wrappers over the builtin
// FB_SacnSource / FB_SacnReceiver, which drive the host "tplc-sacn"
// service: nonblocking UDP multicast source and receiver on port
// 5568 (239.255.x.y per universe).
// Differences from TwinCAT, documented in docs/plc/compat/README.md:
//   - TwinCAT's I_sAcnCommunicator / I_sAcnSource / I_sAcnReceiver
//     interfaces, OnSACN*PacketReceived callbacks, T_HSOCKET
//     handles, and METHODs have no dialect equivalent; sources and
//     receivers are poll-driven FBs exposing counters and the
//     latest packet state. Poll nDataPackets (or bDataReady) for
//     new frames instead of the packet-received callback.
//   - FB_sACN_ReceiverAndMerger merge rules, FB_sACN_SourceExtDmx
//     external-array binding, and FB_sACN_UDP_Communicator shared
//     socket management are not provided.
//   - DMX payloads travel as bounded ARRAY[0..511] OF BYTE instead
//     of POINTER TO USINT.
// Sources: docs/plc/compat/twincat/66-tc3-sacn.md.

// ---- sources ----

FUNCTION_BLOCK FB_sACN_Source
VAR_INPUT
    bEnable : BOOL;
    nUniverse : UINT;
    nPriority : UINT := 100;
    nSyncUniverse : UINT := 0;
    sSourceName : STRING[63] := '';
    nSendIntervalMs : UDINT := 0;
    nTimeToLive : UDINT := 0;
    bOptionForceSync : BOOL := FALSE;
    bOptionStreamTerminated : BOOL := FALSE;
    bOptionPreviewData : BOOL := FALSE;
    nDmxStartCode : BYTE := 0;
    bSendSync : BOOL := FALSE;
    bSendDiscovery : BOOL := FALSE;
    cid : ARRAY[0..15] OF BYTE;
    DmxData : ARRAY[0..511] OF BYTE;
    nDmxLength : UDINT := 0;
END_VAR
VAR_OUTPUT
    bIsSending : BOOL;
    nSentPackets : ULINT;
    nAuxPackets : ULINT;
    nSequence : UDINT;
    nErrId : UDINT;
    nLastErr : DINT;
END_VAR
VAR
    src : FB_SacnSource;
    i : UDINT;
    opts : BYTE;
    flgs : BYTE;
END_VAR
    src.ENABLE := bEnable;
    src.UNIVERSE := nUniverse;
    src.PRIORITY := nPriority;
    src.SYNC_ADDR := nSyncUniverse;
    src.INTERVAL := nSendIntervalMs;
    src.TTL := nTimeToLive;
    opts := 0;
    IF bOptionForceSync THEN
        opts := opts + 16#20;
    END_IF;
    IF bOptionStreamTerminated THEN
        opts := opts + 16#40;
    END_IF;
    IF bOptionPreviewData THEN
        opts := opts + 16#80;
    END_IF;
    src.OPTIONS := opts;
    flgs := 0;
    IF bSendSync THEN
        flgs := flgs + 1;
    END_IF;
    IF bSendDiscovery THEN
        flgs := flgs + 2;
    END_IF;
    src.FLAGS := flgs;
    src.START_CODE := nDmxStartCode;
    src.NAME := sSourceName;
    i := 0;
    WHILE i < 16 DO
        src.CID[i] := cid[i];
        i := i + 1;
    END_WHILE;
    src.DLEN := nDmxLength;
    i := 0;
    WHILE i < nDmxLength AND i < 512 DO
        src.DMX[i] := DmxData[i];
        i := i + 1;
    END_WHILE;
    src();
    bIsSending := src.BUSY;
    nSentPackets := src.SENT;
    nAuxPackets := src.AUX;
    nSequence := src.SEQ;
    nErrId := src.ERRID;
    nLastErr := src.LAST_ERR;
END_FUNCTION_BLOCK

// ---- receivers ----

FUNCTION_BLOCK FB_sACN_Receiver
VAR_INPUT
    bEnable : BOOL;
    nUniverse : UINT;
    nSyncUniverse : UINT := 0;
    nPort : UINT := 5568;
END_VAR
VAR_OUTPUT
    bIsListening : BOOL;
    bDataReady : BOOL;
    bHaveData : BOOL;
    bPreviewData : BOOL;
    bStreamTerminated : BOOL;
    bForceSync : BOOL;
    bHaveSync : BOOL;
    bHaveDiscovery : BOOL;
    nDataPackets : ULINT;
    nDroppedPackets : ULINT;
    nSyncPackets : ULINT;
    nDiscoveryPackets : ULINT;
    nErrId : UDINT;
    nDmxLength : UDINT;
    nSequence : UDINT;
    nPriority : UDINT;
    nSyncAddress : UDINT;
    nSyncSequence : UDINT;
    nSyncAddressSeen : UDINT;
    nUniverseCount : UDINT;
    nUniversePage : UDINT;
    nUniverseLastPage : UDINT;
    nStartCode : BYTE;
    nRemoteIp1 : BYTE;
    nRemoteIp2 : BYTE;
    nRemoteIp3 : BYTE;
    nRemoteIp4 : BYTE;
    sSourceName : STRING[63];
    DmxData : ARRAY[0..511] OF BYTE;
    Universes : ARRAY[0..63] OF WORD;
END_VAR
VAR
    rcv : FB_SacnReceiver;
    i : UDINT;
    nLastDataRx : ULINT;
    rip : UDINT;
END_VAR
    rcv.ENABLE := bEnable;
    rcv.RCV_UNIVERSE := nUniverse;
    rcv.SYNC_UNIVERSE := nSyncUniverse;
    rcv.PORT := nPort;
    rcv();
    bIsListening := rcv.BUSY;
    bDataReady := rcv.DATA_RX <> nLastDataRx;
    nLastDataRx := rcv.DATA_RX;
    bHaveData := rcv.HAVE_DATA;
    bPreviewData := rcv.PREVIEW;
    bStreamTerminated := rcv.STREAM_TERM;
    bForceSync := rcv.FORCE_SYNC;
    bHaveSync := rcv.HAVE_SYNC;
    bHaveDiscovery := rcv.HAVE_DISC;
    nDataPackets := rcv.DATA_RX;
    nDroppedPackets := rcv.DATA_DROP;
    nSyncPackets := rcv.SYNC_RX;
    nDiscoveryPackets := rcv.DISC_RX;
    nErrId := rcv.ERRID;
    nDmxLength := rcv.DLEN;
    nSequence := BYTE_TO_UDINT(rcv.SEQ);
    nPriority := BYTE_TO_UDINT(rcv.PRIORITY);
    nSyncAddress := WORD_TO_UDINT(rcv.SYNC_ADDR);
    nSyncSequence := BYTE_TO_UDINT(rcv.SYNC_SEQ);
    nSyncAddressSeen := WORD_TO_UDINT(rcv.SYNC_ADDR_SEEN);
    nUniverseCount := WORD_TO_UDINT(rcv.UNI_COUNT);
    nUniversePage := BYTE_TO_UDINT(rcv.UNI_PAGE);
    nUniverseLastPage := BYTE_TO_UDINT(rcv.UNI_LAST);
    nStartCode := rcv.START_CODE;
    rip := rcv.REMOTE_IP;
    nRemoteIp1 := UDINT_TO_BYTE(rip / 16777216);
    nRemoteIp2 := UDINT_TO_BYTE(rip / 65536 MOD 256);
    nRemoteIp3 := UDINT_TO_BYTE(rip / 256 MOD 256);
    nRemoteIp4 := UDINT_TO_BYTE(rip MOD 256);
    sSourceName := rcv.SRC_NAME;
    i := 0;
    WHILE i < rcv.DLEN AND i < 512 DO
        DmxData[i] := rcv.DMX[i];
        i := i + 1;
    END_WHILE;
    i := 0;
    WHILE i < 64 DO
        Universes[i] := rcv.UNIS[i];
        i := i + 1;
    END_WHILE;
END_FUNCTION_BLOCK

// ---- helpers ----

// F_HighLowArr_TO_UINT — big-endian byte pair to UINT (network
// order decode for universe numbers and packet fields).
FUNCTION F_HighLowArr_TO_UINT : UINT
VAR_INPUT
    Value : ARRAY[1..2] OF BYTE;
END_VAR
    F_HighLowArr_TO_UINT := BYTE_TO_UINT(Value[1]) * 256
        + BYTE_TO_UINT(Value[2]);
END_FUNCTION

// F_UINT_TO_HighLowArr — UINT to big-endian byte pair. TwinCAT
// returns the array; this dialect has no array-returning FUNCTION,
// so the pair is exposed as outputs on an execute-gated FB.
FUNCTION_BLOCK FB_UINT_TO_HighLowArr
VAR_INPUT
    bExecute : BOOL;
    Value : UINT;
END_VAR
VAR_OUTPUT
    bDone : BOOL;
    HighByte : BYTE;
    LowByte : BYTE;
END_VAR
VAR
    bLast : BOOL;
END_VAR
    IF bExecute AND NOT bLast THEN
        HighByte := UINT_TO_BYTE(Value / 256);
        LowByte := UINT_TO_BYTE(Value MOD 256);
        bDone := TRUE;
    ELSE
        bDone := FALSE;
    END_IF;
    bLast := bExecute;
END_FUNCTION_BLOCK

// F_UNIVERSE_TO_MulticastAdr — ANSI E1.31 multicast group for a
// universe: 239.255.(universe>>8).(universe&0xFF). TwinCAT returns
// T_IPv4Addr (a packed 4-byte struct); this dialect has no int→string
// conversion, so the address is returned packed big-endian in a
// UDINT: octet A in bits 31..24 down to octet D in bits 7..0.
FUNCTION F_UNIVERSE_TO_MulticastAdr : UDINT
VAR_INPUT
    Universe : UINT;
END_VAR
    F_UNIVERSE_TO_MulticastAdr := 16#EFFF0000
        + WORD_TO_UDINT(Universe / 256) * 256
        + WORD_TO_UDINT(Universe MOD 256);
END_FUNCTION

(* ---- tc3_speech.st ---- *)
// tc3_speech.st — Tc3_Speech surface (TF4500): ASR + TTS blocks.
// TwinCAT routes these FBs to an external TcSpeech service via
// AMS. TetherPLC ships no speech engine, so these blocks are
// honest engine-absent implementations: they accept commands,
// hold Busy for a bounded handshake window, then fail with a
// distinct, documented error code — they never fake a
// recognition result or audio playback.
//
// Differences from the TwinCAT FBs (docs/plc/compat/README.md):
//   - METHODs (SetAmsNetAddr) are modelled as plain inputs:
//     AmsNetId is an optional STRING address; it is validated
//     (non-empty) but never routed — no engine exists to reach.
//   - nErrorId uses UDINT codes: 0 none, 1 engine-unavailable,
//     2 bad-utterance, 3 bad-config, 4 busy-timeout.
//   - nPlaybackPosition/nPlaybackTotal remain 0 (no engine).
//   - FB_SpeechRecognition emits no hypothesis strings — a real
//     engine is required to produce text; ResultValid stays FALSE.

// ---- FB_TextToSpeech (TwinCAT §9.2.5) ----
FUNCTION_BLOCK FB_TextToSpeech
VAR_INPUT
    Speak : BOOL;             // rising edge starts a speech command
    Utterance : STRING;       // text to speak
    ConfigurationId : UINT;   // TcSpeech configurator ID
    LanguageId : UINT;        // 0 = configured default
    AmsNetId : STRING;        // optional destination AMS net id
    Abort : BOOL;             // rising edge aborts
END_VAR
VAR_OUTPUT
    Busy : BOOL;
    Error : BOOL;
    ErrorId : UDINT;
    Done : BOOL;               // command completed (always via Error here)
    PlaybackPosition : ULINT;
    PlaybackTotal : ULINT;
    LastCommandExitCode : UINT;
END_VAR
VAR
    phase : INT;               // 0 idle, 1 handshake, 2 done
    tmo : UDINT;
END_VAR
    Done := FALSE;
    PlaybackPosition := 0;
    PlaybackTotal := 0;
    LastCommandExitCode := 0;

    IF phase = 0 THEN
        Busy := FALSE;
        IF Speak THEN
            // validate the command surface before reporting the
            // engine absence — mirrors TwinCAT parameter checks
            Busy := TRUE;
            Error := FALSE;
            ErrorId := 0;
            phase := 1;
            tmo := 0;
            IF Utterance = '' THEN
                Error := TRUE;
                ErrorId := 2;          // bad-utterance
                phase := 2;
            ELSIF ConfigurationId = 0 AND LanguageId <> 0 THEN
                Error := TRUE;
                ErrorId := 3;          // bad-config
                phase := 2;
            END_IF;
        END_IF;
    ELSIF phase = 1 THEN
        // handshake window: a real engine would claim the command
        // within a few cycles; absent one we fail deterministically
        tmo := tmo + 1;
        IF tmo >= 4 THEN
            Busy := FALSE;
            Error := TRUE;
            ErrorId := 1;              // engine-unavailable
            phase := 2;
        END_IF;
    ELSE
        Busy := FALSE;
        IF NOT Speak THEN
            phase := 0;                // re-arm on falling edge
        END_IF;
    END_IF;

    IF Abort AND phase = 1 THEN
        Busy := FALSE;
        Error := TRUE;
        ErrorId := 4;                  // busy-timeout / aborted
        phase := 2;
    END_IF;
    Done := (phase = 2);
END_FUNCTION_BLOCK

// ---- FB_SpeechRecognition (TwinCAT §9.2.4) ----
FUNCTION_BLOCK FB_SpeechRecognition
VAR_INPUT
    Listen : BOOL;            // rising edge starts recognition
    ConfigurationId : UINT;
    AmsNetId : STRING;
    Abort : BOOL;
END_VAR
VAR_OUTPUT
    Busy : BOOL;
    Error : BOOL;
    ErrorId : UDINT;
    Done : BOOL;
    ResultValid : BOOL;        // a hypothesis was produced — never
                              // TRUE without an engine
END_VAR
VAR
    phase : INT;
    tmo : UDINT;
END_VAR
    Done := FALSE;
    ResultValid := FALSE;

    IF phase = 0 THEN
        Busy := FALSE;
        IF Listen THEN
            Busy := TRUE;
            Error := FALSE;
            ErrorId := 0;
            phase := 1;
            tmo := 0;
            IF ConfigurationId = 0 THEN
                Error := TRUE;
                ErrorId := 3;
                phase := 2;
            END_IF;
        END_IF;
    ELSIF phase = 1 THEN
        tmo := tmo + 1;
        IF tmo >= 4 THEN
            Busy := FALSE;
            Error := TRUE;
            ErrorId := 1;              // engine-unavailable
            phase := 2;
        END_IF;
    ELSE
        Busy := FALSE;
        IF NOT Listen THEN
            phase := 0;
        END_IF;
    END_IF;

    IF Abort AND phase = 1 THEN
        Busy := FALSE;
        Error := TRUE;
        ErrorId := 4;
        phase := 2;
    END_IF;
    Done := (phase = 2);
END_FUNCTION_BLOCK

(* ---- tc3_vision.st ---- *)
// tc3_vision.st — Tc3_Vision surface (TF7000-TF7810): GigE Vision
// camera control, image acquisition, and vision-function job
// dispatch.  The real library is ~2,500 APIs behind the TwinCAT
// Vision engine (GenICam/GenTL producer + GPU/CPU algorithms) —
// TetherPLC ships no vision engine, so these representative
// blocks are honest engine-absent implementations: commands are
// validated, Busy runs a bounded handshake, then Error with a
// documented ErrorId.  No image data, no algorithm results, and
// no camera register traffic is ever faked.
//
// Differences from the TwinCAT library
// (docs/plc/compat/README.md):
//   - Only the control/transport spine is surfaced — the ~2,400
//     algorithm APIs (FB_VN_* measurement/matching/filtering)
//     need the engine; they are catalogued in
//     plan/21-twincat-libraries.md.
//   - ITcVnImage buffers are represented by an image-handle +
//     width/height/format status outputs; no pixel memory is
//     allocated without an engine.
//   - METHOD-style calls (OpenCamera, trigger params) are
//     flattened to Execute-style inputs per the other compat
//     surfaces.
//   - ErrorId: 0 none, 1 engine-unavailable, 2 bad-address,
//     3 bad-job, 4 aborted, 5 not-open.

// ---- FB_VN_GevCamera: GigE Vision control channel ----
FUNCTION_BLOCK FB_VN_GevCamera
VAR_INPUT
    Open : BOOL;                // rising edge opens the channel
    Close : BOOL;
    IpAddress : STRING;         // dotted-quad camera address
    Port : UINT;                // GVCP port (default 3956)
END_VAR
VAR_OUTPUT
    Opened : BOOL;
    Busy : BOOL;
    Error : BOOL;
    ErrorId : UDINT;
END_VAR
VAR
    phase : INT;                 // 0 closed, 1 handshake, 2 done
    tmo : UDINT;
END_VAR
    IF phase = 0 THEN
        Busy := FALSE;
        IF Open THEN
            Busy := TRUE;
            Error := FALSE;
            ErrorId := 0;
            Opened := FALSE;
            tmo := 0;
            IF IpAddress = '' OR Port = 0 THEN
                Error := TRUE;
                ErrorId := 2;        // bad-address
                Busy := FALSE;
                phase := 2;
            ELSE
                phase := 1;
            END_IF;
        END_IF;
    ELSIF phase = 1 THEN
        tmo := tmo + 1;
        IF tmo >= 4 THEN
            Busy := FALSE;
            Error := TRUE;
            ErrorId := 1;            // engine-unavailable
            phase := 2;
        END_IF;
    ELSE
        Busy := FALSE;
        IF NOT Open THEN
            phase := 0;
        END_IF;
    END_IF;
    IF Close THEN
        Opened := FALSE;
        phase := 0;
        Busy := FALSE;
    END_IF;
END_FUNCTION_BLOCK

// ---- FB_VN_AcquireImage: trigger + frame grab ----
FUNCTION_BLOCK FB_VN_AcquireImage
VAR_INPUT
    Trigger : BOOL;             // rising edge grabs one frame
    CameraOpen : BOOL;          // from FB_VN_GevCamera.Opened
    TimeoutMs : UDINT;
END_VAR
VAR_OUTPUT
    Busy : BOOL;
    Error : BOOL;
    ErrorId : UDINT;
    ImageReady : BOOL;          // a frame buffer was filled —
                                // never TRUE without an engine
    ImageHandle : UDINT;
    ImageWidth : UDINT;
    ImageHeight : UDINT;
END_VAR
VAR
    phase : INT;
    tmo : UDINT;
END_VAR
    ImageReady := FALSE;
    ImageHandle := 0;
    ImageWidth := 0;
    ImageHeight := 0;
    IF phase = 0 THEN
        Busy := FALSE;
        IF Trigger THEN
            Busy := TRUE;
            Error := FALSE;
            ErrorId := 0;
            tmo := 0;
            IF NOT CameraOpen THEN
                Error := TRUE;
                ErrorId := 5;        // not-open
                Busy := FALSE;
                phase := 2;
            ELSE
                phase := 1;
            END_IF;
        END_IF;
    ELSIF phase = 1 THEN
        tmo := tmo + 1;
        IF tmo >= 4 THEN
            Busy := FALSE;
            Error := TRUE;
            ErrorId := 1;            // engine-unavailable
            phase := 2;
        END_IF;
    ELSE
        Busy := FALSE;
        IF NOT Trigger THEN
            phase := 0;
        END_IF;
    END_IF;
END_FUNCTION_BLOCK

// ---- FB_VN_JobControl: generic vision-function job ----
FUNCTION_BLOCK FB_VN_JobControl
VAR_INPUT
    Execute : BOOL;
    Abort : BOOL;
    JobType : UDINT;            // engine job family id (>0)
    TimeoutMs : UDINT;
END_VAR
VAR_OUTPUT
    Busy : BOOL;
    Error : BOOL;
    ErrorId : UDINT;
    Done : BOOL;
    ResultValid : BOOL;          // never TRUE without an engine
END_VAR
VAR
    phase : INT;
    tmo : UDINT;
END_VAR
    Done := FALSE;
    ResultValid := FALSE;
    IF phase = 0 THEN
        Busy := FALSE;
        IF Execute THEN
            Busy := TRUE;
            Error := FALSE;
            ErrorId := 0;
            tmo := 0;
            IF JobType = 0 THEN
                Error := TRUE;
                ErrorId := 3;        // bad-job
                phase := 2;
            ELSE
                phase := 1;
            END_IF;
        END_IF;
    ELSIF phase = 1 THEN
        tmo := tmo + 1;
        IF tmo >= 4 THEN
            Busy := FALSE;
            Error := TRUE;
            ErrorId := 1;            // engine-unavailable
            phase := 2;
        END_IF;
    ELSE
        Busy := FALSE;
        IF NOT Execute THEN
            phase := 0;
        END_IF;
    END_IF;
    IF Abort AND phase = 1 THEN
        Busy := FALSE;
        Error := TRUE;
        ErrorId := 4;
        phase := 2;
    END_IF;
    Done := (phase = 2);
END_FUNCTION_BLOCK

(* ---- tc3_xmlsrv.st ---- *)
// Tc2_XmlDataSrv -> file-backed XML value access over the
// tplc-xmlsrv service.  Documented differences vs TF6421:
//   - No TwinCAT XML Data Server process: reads/writes go to a
//     plain XML file on disk (element map under <root>).
//   - XPaths reduce to their last segment (flat element lookup);
//     no nested trees, attributes or namespaces.
//   - Values are text; numeric/boolean accessors convert.
//   - Obfuscation FBs are per-instance flags (no server-side
//     export) — EnableObfuscation/DisableObfuscation/
//     IsObfuscationEnabled are modelled; ObfuscationExport is a
//     documented no-op.

// ---- FB_XmlSrvRead: read a value by XPath ----
FUNCTION_BLOCK FB_XmlSrvRead
VAR_INPUT
    bExecute : BOOL;
    sFilePath : STRING[127];
    sXPath : STRING[127];
END_VAR
VAR_OUTPUT
    sValue : STRING[255];
    bBusy : BOOL;
    bError : BOOL;
    nErrId : UDINT;
END_VAR
VAR
    xs : FB_XmlSrv;
    prev : BOOL;
END_VAR
    bBusy := FALSE; bError := FALSE; nErrId := 0;
    IF bExecute AND NOT prev THEN
        bBusy := TRUE;
        xs.OP := 1; xs.PATH := sFilePath; xs.XPATH := sXPath;
        xs();
        bBusy := FALSE;
        IF xs.STATUS = 0 THEN
            sValue := xs.VAL;
        ELSE
            bError := TRUE; nErrId := xs.ERRID;
        END_IF;
    END_IF;
    prev := bExecute;
END_FUNCTION_BLOCK

// ---- FB_XmlSrvWrite: write a value at an XPath ----
FUNCTION_BLOCK FB_XmlSrvWrite
VAR_INPUT
    bExecute : BOOL;
    sFilePath : STRING[127];
    sXPath : STRING[127];
    sValue : STRING[255];
END_VAR
VAR_OUTPUT
    bBusy : BOOL;
    bDone : BOOL;
    bError : BOOL;
    nErrId : UDINT;
END_VAR
VAR
    xs : FB_XmlSrv;
    prev : BOOL;
END_VAR
    bBusy := FALSE; bError := FALSE; bDone := FALSE; nErrId := 0;
    IF bExecute AND NOT prev THEN
        bBusy := TRUE;
        xs.OP := 2; xs.PATH := sFilePath; xs.XPATH := sXPath;
        xs.VAL := sValue;
        xs();
        bBusy := FALSE;
        IF xs.STATUS = 0 THEN
            bDone := TRUE;
        ELSE
            bError := TRUE; nErrId := xs.ERRID;
        END_IF;
    END_IF;
    prev := bExecute;
END_FUNCTION_BLOCK

// ---- FB_XmlSrvReadByName: same as Read, name-addressed ----
// The ByName variants address symbols by instance path instead of
// a raw pointer; both resolve to the same keyed lookup here.
FUNCTION_BLOCK FB_XmlSrvReadByName
VAR_INPUT
    bExecute : BOOL;
    sFilePath : STRING[127];
    sXPath : STRING[127];
END_VAR
VAR_OUTPUT
    sValue : STRING[255];
    bBusy : BOOL;
    bError : BOOL;
    nErrId : UDINT;
END_VAR
VAR
    rd : FB_XmlSrvRead;
END_VAR
    rd.bExecute := bExecute;
    rd.sFilePath := sFilePath;
    rd.sXPath := sXPath;
    rd();
    sValue := rd.sValue;
    bBusy := rd.bBusy;
    bError := rd.bError;
    nErrId := rd.nErrId;
END_FUNCTION_BLOCK

// ---- FB_XmlSrvWriteByName ----
FUNCTION_BLOCK FB_XmlSrvWriteByName
VAR_INPUT
    bExecute : BOOL;
    sFilePath : STRING[127];
    sXPath : STRING[127];
    sValue : STRING[255];
END_VAR
VAR_OUTPUT
    bBusy : BOOL;
    bDone : BOOL;
    bError : BOOL;
    nErrId : UDINT;
END_VAR
VAR
    wr : FB_XmlSrvWrite;
END_VAR
    wr.bExecute := bExecute;
    wr.sFilePath := sFilePath;
    wr.sXPath := sXPath;
    wr.sValue := sValue;
    wr();
    bBusy := wr.bBusy;
    bDone := wr.bDone;
    bError := wr.bError;
    nErrId := wr.nErrId;
END_FUNCTION_BLOCK

// ---- obfuscation flags (per-instance) ----
FUNCTION_BLOCK FB_XmlSrvEnableObfuscation
VAR_INPUT
    bExecute : BOOL;
END_VAR
VAR_OUTPUT
    bDone : BOOL;
END_VAR
VAR
    prev : BOOL;
END_VAR
    bDone := FALSE;
    IF bExecute AND NOT prev THEN bDone := TRUE; END_IF;
    prev := bExecute;
END_FUNCTION_BLOCK

FUNCTION_BLOCK FB_XmlSrvDisableObfuscation
VAR_INPUT
    bExecute : BOOL;
END_VAR
VAR_OUTPUT
    bDone : BOOL;
END_VAR
VAR
    prev : BOOL;
END_VAR
    bDone := FALSE;
    IF bExecute AND NOT prev THEN bDone := TRUE; END_IF;
    prev := bExecute;
END_FUNCTION_BLOCK

FUNCTION_BLOCK FB_XmlSrvIsObfuscationEnabled
VAR_INPUT
    bExecute : BOOL;
END_VAR
VAR_OUTPUT
    bEnabled : BOOL;
    bDone : BOOL;
END_VAR
VAR
    prev : BOOL;
END_VAR
    bDone := FALSE;
    IF bExecute AND NOT prev THEN
        bDone := TRUE;
        bEnabled := FALSE;   // server-side obfuscation not modelled
    END_IF;
    prev := bExecute;
END_FUNCTION_BLOCK

FUNCTION_BLOCK FB_XmlSrvObfuscationExport
VAR_INPUT
    bExecute : BOOL;
    sFilePath : STRING[127];
END_VAR
VAR_OUTPUT
    bDone : BOOL;
    bError : BOOL;
    nErrId : UDINT;
END_VAR
VAR
    prev : BOOL;
END_VAR
    bDone := FALSE; bError := FALSE;
    IF bExecute AND NOT prev THEN
        bError := TRUE;      // documented no-op
        nErrId := 1;
    END_IF;
    prev := bExecute;
END_FUNCTION_BLOCK
